(* IEC 61131-3 sources: guidance-for-physical-ai-production-designer-on-aws/source/plan2cell/examples/welding_cell_2_small/plc/trust/robot2/src, 20 files *)

(* ---- E_PlayerState.st ---- *)
(*
 * E_PlayerState
 * States of FB_ProgramPlayer (robot side of the bt2plc zone protocol).
 * Device simulator R2 (robot2), cell welding_cell_2_small. Generated by bt2plc 0.1.0.
 *)

TYPE E_PlayerState :
(
    PS_IDLE         := 0,    (* No program, pose held *)
    PS_NEXT_OP      := 10,   (* Advance to the next op: wStep := k, REQUEST := mask *)
    PS_WAIT_GRANT   := 20,   (* Wait (GRANT AND mask) = mask *)
    PS_DELAY        := 30,   (* Start delay of the op *)
    PS_MOVE         := 40,   (* Trajectory / blind home move *)
    PS_HOLD         := 50,   (* Hold at the end pose *)
    PS_WAIT_RELEASE := 60,   (* REQUEST := 0, wait (GRANT AND mask) = 0 *)
    PS_DONE         := 90,   (* Program finished *)
    PS_ERROR        := 99    (* Program aborted with an error *)
);
END_TYPE

(* ---- E_ProgramState.st ---- *)
(*
 * E_ProgramState
 * VW VASS standard - robot program states.
 * Device simulator R2 (robot2), cell welding_cell_2_small. Generated by bt2plc 0.1.0.
 *)

TYPE E_ProgramState :
(
    PRG_IDLE     := 0,
    PRG_RUNNING  := 1,
    PRG_STOPPED  := 2,
    PRG_PAUSED   := 3,
    PRG_FINISHED := 4,
    PRG_ERROR    := 5
);
END_TYPE

(* ---- E_RobotMode.st ---- *)
(*
 * E_RobotMode
 * VW VASS standard - KUKA KR C4 robot operating modes.
 * Device simulator R2 (robot2), cell welding_cell_2_small. Generated by bt2plc 0.1.0.
 *)

TYPE E_RobotMode :
(
    MODE_UNKNOWN := 0,
    MODE_T1      := 1,       (* Test mode 1 - reduced speed *)
    MODE_T2      := 2,       (* Test mode 2 - programmed speed *)
    MODE_AUT     := 3,       (* Automatic mode *)
    MODE_EXT     := 4        (* External automatic - PLC controlled *)
);
END_TYPE

(* ---- ST_OpDef.st ---- *)
(*
 * ST_OpDef
 * One op of the bt2plc robot program (row of GVL_Program.aOps).
 * Op k plays waypoints GVL_Program.aWp[nFirstWp..nLastWp] under the zone mask dwZoneMask.
 * Blind home op: bBlindHome = TRUE, nFirstWp = nLastWp = 0 (joint move to arHomeDeg over R_HOME_S).
 * Device simulator R2 (robot2), cell welding_cell_2_small. Generated by bt2plc 0.1.0.
 *)

TYPE ST_OpDef :
STRUCT
    sName           : STRING(32);   (* Operation id, e.g. 'W01' *)
    nFirstWp        : INT;          (* First waypoint index in aWp (0 = none) *)
    nLastWp         : INT;          (* Last waypoint index in aWp (0 = none) *)
    dwZoneMask      : DWORD;        (* REQUEST/GRANT bits (zones 0..30, bit 31 = permit) *)
    tDelay          : TIME;         (* Start delay after the grant *)
    tHold           : TIME;         (* Hold time at the end pose *)
    rDelay_s        : REAL;         (* Start delay in s (used by FB_ProgramPlayer) *)
    rHold_s         : REAL;         (* Hold time in s (used by FB_ProgramPlayer) *)
    rVelScale       : REAL;         (* Velocity scale of the trajectory (1.0 = nominal) *)
    bBlindHome      : BOOL;         (* TRUE = blind joint move to the home pose *)
END_STRUCT
END_TYPE

(* ---- ST_PROFIsafe_Trailer.st ---- *)
(*
 * ST_PROFIsafe_Trailer
 * PROFIsafe trailer - 4 bytes appended by the safety layer (status + 3-byte CRC).
 * Device simulator R2 (robot2), cell welding_cell_2_small. Generated by bt2plc 0.1.0.
 *)

TYPE ST_PROFIsafe_Trailer :
STRUCT
    byStatus        : BYTE;                     (* Status/Control byte *)
    abyCRC          : ARRAY[0..2] OF BYTE;      (* 3-byte CRC *)
END_STRUCT
END_TYPE

(* ---- ST_SafeInput.st ---- *)
(*
 * ST_SafeInput
 * PROFIsafe (Slot 1 - FDIO64) safe inputs: robot -> PLC, 8 bytes user data.
 * GSDML: 8x Unsigned8 Input + F_MessageTrailer4Byte.
 * Device simulator R2 (robot2), cell welding_cell_2_small. Generated by bt2plc 0.1.0.
 *)

TYPE ST_SafeInput :
STRUCT
    (* Byte 0: Safe robot status *)
    bSafe_DrivesOK          : BOOL;   (* Bit 0: Safe drives monitoring OK *)
    bSafe_RobotStopped      : BOOL;   (* Bit 1: Robot safely stopped (SOS/SS1) *)
    bSafe_ReducedSpeed      : BOOL;   (* Bit 2: Safe reduced speed active (SLS) *)
    bSafe_AxisMonitoring    : BOOL;   (* Bit 3: Safe axis range monitoring OK *)
    bSafe_ToolOK            : BOOL;   (* Bit 4: Safe tool monitoring OK *)
    bSafe_WorkspaceOK       : BOOL;   (* Bit 5: Safe workspace monitoring OK *)
    bSafe_Reserved06        : BOOL;   (* Bit 6: Reserved *)
    bSafe_Reserved07        : BOOL;   (* Bit 7: Reserved *)

    (* Byte 1: Safe gate/zone status *)
    bSafe_Gate1Closed       : BOOL;   (* Bit 0: Safety gate 1 closed *)
    bSafe_Gate2Closed       : BOOL;   (* Bit 1: Safety gate 2 closed *)
    bSafe_Gate3Closed       : BOOL;   (* Bit 2: Safety gate 3 closed *)
    bSafe_LightCurtainOK    : BOOL;   (* Bit 3: Light curtain free *)
    bSafe_EStopOK           : BOOL;   (* Bit 4: E-Stop not pressed (NC) *)
    bSafe_EnablingDevice    : BOOL;   (* Bit 5: Enabling device pressed (T1/T2) *)
    bSafe_OperatorSafe      : BOOL;   (* Bit 6: Operator protection OK *)
    bSafe_Reserved17        : BOOL;   (* Bit 7: Reserved *)

    (* Byte 2: Extended safe status *)
    bSafe_STO_Active        : BOOL;   (* Bit 0: Safe Torque Off active *)
    bSafe_SS1_Active        : BOOL;   (* Bit 1: Safe Stop 1 active *)
    bSafe_SS2_Active        : BOOL;   (* Bit 2: Safe Stop 2 active *)
    bSafe_SOS_Active        : BOOL;   (* Bit 3: Safe Operating Stop active *)
    bSafe_SLS_Active        : BOOL;   (* Bit 4: Safely-Limited Speed active *)
    bSafe_SLP_Active        : BOOL;   (* Bit 5: Safely-Limited Position active *)
    bSafe_Reserved26        : BOOL;   (* Bit 6: Reserved *)
    bSafe_FaultPresent      : BOOL;   (* Bit 7: Safety fault present *)

    (* Bytes 3-7: Additional safe signals *)
    bySafe_UserInput3       : BYTE;   (* Byte 3: User safe input *)
    bySafe_UserInput4       : BYTE;   (* Byte 4: User safe input *)
    bySafe_UserInput5       : BYTE;   (* Byte 5: User safe input *)
    bySafe_UserInput6       : BYTE;   (* Byte 6: User safe input *)
    bySafe_UserInput7       : BYTE;   (* Byte 7: User safe input *)
END_STRUCT
END_TYPE

(* ---- ST_SafeOutput.st ---- *)
(*
 * ST_SafeOutput
 * PROFIsafe (Slot 1 - FDIO64) safe outputs: PLC -> robot, 8 bytes user data.
 * GSDML: 8x Unsigned8 Output + F_MessageTrailer4Byte.
 * Device simulator R2 (robot2), cell welding_cell_2_small. Generated by bt2plc 0.1.0.
 *)

TYPE ST_SafeOutput :
STRUCT
    (* Byte 0: Safe control from PLC *)
    bSafe_DriveEnable       : BOOL;   (* Bit 0: Enable drives (safe channel) *)
    bSafe_ExternalEStop     : BOOL;   (* Bit 1: External E-Stop request *)
    bSafe_SafeStop1         : BOOL;   (* Bit 2: Request Safe Stop 1 *)
    bSafe_SafeStop2         : BOOL;   (* Bit 3: Request Safe Stop 2 *)
    bSafe_ReducedSpeedReq   : BOOL;   (* Bit 4: Request safe reduced speed *)
    bSafe_GateOverride      : BOOL;   (* Bit 5: Gate override (maintenance) *)
    bSafe_Reserved06        : BOOL;   (* Bit 6: Reserved *)
    bSafe_Reserved07        : BOOL;   (* Bit 7: Reserved *)

    (* Byte 1: Safe zone control *)
    bSafe_Zone1Enable       : BOOL;   (* Bit 0: Enable workspace zone 1 *)
    bSafe_Zone2Enable       : BOOL;   (* Bit 1: Enable workspace zone 2 *)
    bSafe_Zone3Enable       : BOOL;   (* Bit 2: Enable workspace zone 3 *)
    bSafe_Zone4Enable       : BOOL;   (* Bit 3: Enable workspace zone 4 *)
    bSafe_Reserved14        : BOOL;   (* Bit 4: Reserved *)
    bSafe_Reserved15        : BOOL;   (* Bit 5: Reserved *)
    bSafe_Reserved16        : BOOL;   (* Bit 6: Reserved *)
    bSafe_Reserved17        : BOOL;   (* Bit 7: Reserved *)

    (* Bytes 2-7: Additional safe control *)
    bySafe_UserOutput2      : BYTE;   (* Byte 2: User safe output *)
    bySafe_UserOutput3      : BYTE;   (* Byte 3: User safe output *)
    bySafe_UserOutput4      : BYTE;   (* Byte 4: User safe output *)
    bySafe_UserOutput5      : BYTE;   (* Byte 5: User safe output *)
    bySafe_UserOutput6      : BYTE;   (* Byte 6: User safe output *)
    bySafe_UserOutput7      : BYTE;   (* Byte 7: User safe output *)
END_STRUCT
END_TYPE

(* ---- ST_VASS_ControlWord.st ---- *)
(*
 * ST_VASS_ControlWord
 * VASS PLC control word - output bytes 0-1 (PLC -> robot), Slot 2 DIO256.
 * Device simulator R2 (robot2), cell welding_cell_2_small. Generated by bt2plc 0.1.0.
 *)

TYPE ST_VASS_ControlWord :
STRUCT
    (* Byte 0 *)
    bDrivesOn           : BOOL;   (* Bit 0: Enable drives *)
    bProgStart          : BOOL;   (* Bit 1: Start program *)
    bProgStop           : BOOL;   (* Bit 2: Stop program *)
    bProgCancel         : BOOL;   (* Bit 3: Cancel program *)
    bModeRequest        : BOOL;   (* Bit 4: Request EXT mode *)
    bReset              : BOOL;   (* Bit 5: Reset error *)
    bHomeRequest        : BOOL;   (* Bit 6: Move to home *)
    bConfirm            : BOOL;   (* Bit 7: Confirm/acknowledge *)

    (* Byte 1 *)
    bJobRequest         : BOOL;   (* Bit 8: New job request *)
    bGripperOpen        : BOOL;   (* Bit 9: Open gripper *)
    bGripperClose       : BOOL;   (* Bit 10: Close gripper *)
    bPeriphRelease      : BOOL;   (* Bit 11: Release peripheral *)
    bSpeedOverride      : BOOL;   (* Bit 12: Apply speed override *)
    bReserved13         : BOOL;   (* Bit 13: Reserved *)
    bReserved14         : BOOL;   (* Bit 14: Reserved *)
    bReserved15         : BOOL;   (* Bit 15: Reserved *)
END_STRUCT
END_TYPE

(* ---- ST_VASS_InputTelegram.st ---- *)
(*
 * ST_VASS_InputTelegram
 * Full VASS input telegram - 32 bytes (robot -> PLC), Slot 2 DIO256 inputs.
 * bt2plc use: bytes 4-5 wCurrentStep = op index (GVL_Program.STEP_BYTE),
 *             bytes 16-27 joint angles A1..A6 (FB_JointAngleEncoder),
 *             bytes 28-31 zone REQUEST DWORD LE (GVL_Program.REQ_BYTE).
 * Device simulator R2 (robot2), cell welding_cell_2_small. Generated by bt2plc 0.1.0.
 *)

TYPE ST_VASS_InputTelegram :
STRUCT
    stStatusWord        : ST_VASS_StatusWord;     (* Bytes 0-1:   Status word *)
    wActiveJobNr        : WORD;                   (* Bytes 2-3:   Active job number *)
    wCurrentStep        : WORD;                   (* Bytes 4-5:   Current program step *)
    wSpeedActual        : WORD;                   (* Bytes 6-7:   Actual speed % *)
    wActiveToolNr       : WORD;                   (* Bytes 8-9:   Active tool number *)
    wErrorCode          : WORD;                   (* Bytes 10-11: Active error code *)
    wWarningCode        : WORD;                   (* Bytes 12-13: Active warning code *)
    wPositionX          : INT;                    (* Bytes 14-15: Position X (0.1mm) *)
    wPositionY          : INT;                    (* Bytes 16-17: Position Y (0.1mm) *)
    wPositionZ          : INT;                    (* Bytes 18-19: Position Z (0.1mm) *)
    wUserWord10         : WORD;                   (* Bytes 20-21: User data *)
    wUserWord11         : WORD;                   (* Bytes 22-23: User data *)
    wUserWord12         : WORD;                   (* Bytes 24-25: User data *)
    wUserWord13         : WORD;                   (* Bytes 26-27: User data *)
    wUserWord14         : WORD;                   (* Bytes 28-29: User data *)
    wUserWord15         : WORD;                   (* Bytes 30-31: User data *)
END_STRUCT
END_TYPE

(* ---- ST_VASS_OutputTelegram.st ---- *)
(*
 * ST_VASS_OutputTelegram
 * Full VASS output telegram - 32 bytes (PLC -> robot), Slot 2 DIO256 outputs.
 * bt2plc use: bytes 4-5 PLAN_ID WORD LE during a production job (GVL_Program.PLAN_ID_BYTE),
 *             bytes 12-15 zone GRANT DWORD LE (GVL_Program.GRANT_BYTE).
 * Device simulator R2 (robot2), cell welding_cell_2_small. Generated by bt2plc 0.1.0.
 *)

TYPE ST_VASS_OutputTelegram :
STRUCT
    stControlWord       : ST_VASS_ControlWord;    (* Bytes 0-1:   Control word *)
    wJobNr              : WORD;                   (* Bytes 2-3:   Requested job number *)
    wParameter1         : WORD;                   (* Bytes 4-5:   Parameter 1 *)
    wParameter2         : WORD;                   (* Bytes 6-7:   Parameter 2 *)
    wSpeedOverride      : WORD;                   (* Bytes 8-9:   Speed override % *)
    wToolRequest        : WORD;                   (* Bytes 10-11: Tool change request *)
    wUserWord6          : WORD;                   (* Bytes 12-13: User command data *)
    wUserWord7          : WORD;                   (* Bytes 14-15: User command data *)
    wUserWord8          : WORD;                   (* Bytes 16-17: User command data *)
    wUserWord9          : WORD;                   (* Bytes 18-19: User command data *)
    wUserWord10         : WORD;                   (* Bytes 20-21: User command data *)
    wUserWord11         : WORD;                   (* Bytes 22-23: User command data *)
    wUserWord12         : WORD;                   (* Bytes 24-25: User command data *)
    wUserWord13         : WORD;                   (* Bytes 26-27: User command data *)
    wUserWord14         : WORD;                   (* Bytes 28-29: User command data *)
    wUserWord15         : WORD;                   (* Bytes 30-31: User command data *)
END_STRUCT
END_TYPE

(* ---- ST_VASS_StatusWord.st ---- *)
(*
 * ST_VASS_StatusWord
 * VASS robot status word - input bytes 0-1 (robot -> PLC), Slot 2 DIO256.
 * Device simulator R2 (robot2), cell welding_cell_2_small. Generated by bt2plc 0.1.0.
 *)

TYPE ST_VASS_StatusWord :
STRUCT
    (* Byte 0 *)
    bDrivesPowered      : BOOL;   (* Bit 0: Drives are powered on *)
    bProgRunning        : BOOL;   (* Bit 1: Program is running *)
    bAtHome             : BOOL;   (* Bit 2: Robot at home position *)
    bInPosition         : BOOL;   (* Bit 3: Robot in target position *)
    bModeExt            : BOOL;   (* Bit 4: External automatic mode active *)
    bReady              : BOOL;   (* Bit 5: Robot ready for command *)
    bError              : BOOL;   (* Bit 6: Error present *)
    bWarning            : BOOL;   (* Bit 7: Warning present *)

    (* Byte 1 *)
    bSafetyGateOK       : BOOL;   (* Bit 8: Safety gate closed *)
    bEStopNotActive     : BOOL;   (* Bit 9: E-Stop NOT active (NC logic) *)
    bProgFinished       : BOOL;   (* Bit 10: Program/job finished *)
    bJobAcknowledge     : BOOL;   (* Bit 11: Job number acknowledged *)
    bToolActive         : BOOL;   (* Bit 12: Tool/gripper active *)
    bPartPresent        : BOOL;   (* Bit 13: Part present in gripper *)
    bPeriphReady        : BOOL;   (* Bit 14: Peripheral devices ready *)
    bMaintRequired      : BOOL;   (* Bit 15: Maintenance required *)
END_STRUCT
END_TYPE

(* ---- ST_Waypoint.st ---- *)
(*
 * ST_Waypoint
 * One trajectory waypoint (row of GVL_Program.aWp). Flat fields for portability.
 * rT = seconds from op start; angles in degrees (KUKA A1..A6 after joint sign/offset mapping).
 * Device simulator R2 (robot2), cell welding_cell_2_small. Generated by bt2plc 0.1.0.
 *)

TYPE ST_Waypoint :
STRUCT
    rT              : REAL;         (* Time from op start (s) *)
    rA1             : REAL;         (* Axis 1 (deg) *)
    rA2             : REAL;         (* Axis 2 (deg) *)
    rA3             : REAL;         (* Axis 3 (deg) *)
    rA4             : REAL;         (* Axis 4 (deg) *)
    rA5             : REAL;         (* Axis 5 (deg) *)
    rA6             : REAL;         (* Axis 6 (deg) *)
END_STRUCT
END_TYPE

(* ---- GVL_DeviceParams.st ---- *)
NAMESPACE GVL_DeviceParams
(*
 * GVL_DeviceParams
 * PROFINET device identity parameters.
 * Device simulator R2 (robot2, station kuka-robi2), cell welding_cell_2_small. Generated by bt2plc 0.1.0.
 *
 * These parameters configure how the CODESYS PROFINET Device presents itself
 * on the network. They MUST match what the Siemens PLC expects (from the GSDML).
 *
 * In CODESYS, these are typically set via:
 *   1. The "PROFINET Device IEC Objects" tab in the device editor
 *   2. Or programmatically by writing to the device parameter structure
 *
 * The CODESYS PROFINET Device stack reads these at startup and uses them
 * in DCP responses and during the PROFINET connection establishment.
 *
 * IMPORTANT: The default CODESYS values (VendorId=0x02CC, DeviceId=0x1017)
 * will NOT work with the Siemens PLC that expects KUKA (0x019B / 0x0301).
 * You MUST override them.
 *)

{attribute 'qualified_only'}
VAR_GLOBAL
    (* === KUKA VKRCnexxt Device Identity === *)
    (* These values come from GSDML-V2.25-KUKA-Roboter-GmbH-VKR C4-Device-V1.0 *)

    VENDOR_ID           : UINT        := 16#019B;                 (* KUKA Roboter GmbH *)
    DEVICE_ID           : UINT        := 16#0301;                 (* VKR C4 Device *)
    STATION_TYPE        : STRING(240) := 'KUKA VKR C4';           (* Station type string *)
    DEVICE_TYPE         : STRING(28)  := 'KUKA VKR C4';           (* Device type string *)
    ORDER_ID            : STRING(20)  := 'KUKA VKRC nexxt';       (* Order number *)
    HW_REVISION         : UINT        := 1;                       (* Hardware revision *)
    SW_REV_PREFIX       : USINT       := 16#56;                   (* 'V' in ASCII *)
    SW_REV_MAJOR        : UINT        := 8;                       (* V8.x *)
    SW_REV_MINOR        : UINT        := 2;                       (* x.2 *)
    SW_REV_PATCH        : UINT        := 0;                       (* x.x.0 *)

    (* === Module Identification Numbers (from GSDML) === *)
    MODULE_IDENT_DAP    : DWORD       := DWORD#16#00000301;       (* DAP - Slot 0 *)
    MODULE_IDENT_FDIO64 : DWORD       := DWORD#16#0000008F;       (* PROFIsafe - Slot 1 *)
    MODULE_IDENT_DIO256 : DWORD       := DWORD#16#00001000;       (* VASS telegram - Slot 2 *)
    SUBMODULE_IDENT     : DWORD       := DWORD#16#00000001;       (* Submodule ident (all slots) *)

    (* === PROFIsafe Parameters (Slot 1) === *)
    (* These must match the F-parameter record in the PLC safety configuration *)
    F_SIL_LEVEL         : UINT        := 3;                       (* SIL 3 *)
    F_CRC_LENGTH        : UINT        := 3;                       (* 3-byte CRC *)
    F_WD_TIME_DEFAULT   : UINT        := 500;                     (* Watchdog 500ms *)
    F_BLOCK_ID          : UINT        := 0;                       (* Block ID *)
    F_PAR_CRC_DEFAULT   : UINT        := 16#FF59;                 (* Default F_Par_CRC = 65369 *)
END_VAR
END_NAMESPACE

(* ---- GVL_IO.st ---- *)
NAMESPACE GVL_IO
(*
 * GVL_IO
 * Global variable list for the PROFINET device I/O mapping.
 * Device simulator R2 (robot2, station kuka-robi2), cell welding_cell_2_small. Generated by bt2plc 0.1.0.
 *
 * These variables are mapped to the PROFINET device modules via the I/O Mapping tab.
 * Do NOT use AT addresses - the mapping is done in the device configuration.
 * Only PLC_PRG accesses this GVL: it copies the commands into local images and writes
 * the robot status back as a whole array / as scalars (the FBs never touch GVL_IO).
 *
 * Module mapping (set in I/O Mapping tab of each module):
 *   SafeIO_FDIO64 (Slot 1):
 *     "8 safe digital inputs" channels  -> GVL_IO.bySafeIn0..bySafeIn7
 *     "8 safe digital outputs" channels -> GVL_IO.bySafeOut0..bySafeOut7
 *
 *   VASS_DIO256 (Slot 2):
 *     Input channel  -> GVL_IO.aVassInputData
 *     Output channel -> GVL_IO.aVassOutputData
 *)

{attribute 'qualified_only'}
VAR_GLOBAL
    (* ========================================================================
       SLOT 1 - PROFIsafe FDIO64 Module
       8 individual USINT/BYTE channels per direction
       Map each one to the corresponding "8 safe digital inputs/outputs" row
       ======================================================================== *)

    (* Safe Inputs: Robot -> PLC (mapped to "8 safe digital inputs" channels) *)
    bySafeIn0       : BYTE;     (* Safe input byte 0: Drive status *)
    bySafeIn1       : BYTE;     (* Safe input byte 1: Gate/protection *)
    bySafeIn2       : BYTE;     (* Safe input byte 2: STO/SS1/SS2/SOS/SLS *)
    bySafeIn3       : BYTE;     (* Safe input byte 3: User *)
    bySafeIn4       : BYTE;     (* Safe input byte 4: User *)
    bySafeIn5       : BYTE;     (* Safe input byte 5: User *)
    bySafeIn6       : BYTE;     (* Safe input byte 6: User *)
    bySafeIn7       : BYTE;     (* Safe input byte 7: User *)

    (* Safe Outputs: PLC -> Robot (mapped to "8 safe digital outputs" channels) *)
    bySafeOut0      : BYTE;     (* Safe output byte 0: Drive enable, E-Stop, SS1/SS2 *)
    bySafeOut1      : BYTE;     (* Safe output byte 1: Zone enables *)
    bySafeOut2      : BYTE;     (* Safe output byte 2: User *)
    bySafeOut3      : BYTE;     (* Safe output byte 3: User *)
    bySafeOut4      : BYTE;     (* Safe output byte 4: User *)
    bySafeOut5      : BYTE;     (* Safe output byte 5: User *)
    bySafeOut6      : BYTE;     (* Safe output byte 6: User *)
    bySafeOut7      : BYTE;     (* Safe output byte 7: User *)

    (* ========================================================================
       SLOT 2 - DIO256 VASS Telegram
       32 bytes per direction as arrays
       ======================================================================== *)

    (* VASS Inputs: Robot -> PLC (32 bytes) *)
    aVassInputData      : ARRAY[0..31] OF BYTE;

    (* VASS Outputs: PLC -> Robot (32 bytes) *)
    aVassOutputData     : ARRAY[0..31] OF BYTE;
END_VAR
END_NAMESPACE

(* ---- GVL_Program.st ---- *)
NAMESPACE GVL_Program
(*
 * GVL_Program - generated by bt2plc 0.1.0 - DO NOT EDIT
 * Robot program of robot2 (R2) for plan bt_1790934549_welding_cell_2_small (cell welding_cell_2_small)
 * Angles in degrees (KUKA A1..A6 after joint sign/offset), times in seconds from op start.
 *)
{attribute 'qualified_only'}
VAR_GLOBAL
    (* ========================================================================
       IDENTITY / PROTOCOL
       ======================================================================== *)
    ROBOT_TAG               : STRING(16) := 'R2';
    ROBOT_NS                : STRING(32) := 'robot2';
    ROBOT_INDEX             : WORD := WORD#2;
    PLAN_ID                 : WORD := WORD#16#F77E;             (* must match the head PLC *)
    PROD_FOLGE              : WORD := WORD#11;
    HOME_FOLGE              : WORD := WORD#125;
    JOB_NUMBER_BYTE         : BOOL := FALSE;
    STEP_BYTE               : INT := 4;
    REQ_BYTE                : INT := 28;
    GRANT_BYTE              : INT := 12;
    PLAN_ID_BYTE            : INT := 4;
    R_TASK_S                : REAL := 0.0200;                   (* device MainTask interval *)
    R_HOME_S                : REAL := 7.0000;                   (* blind home duration *)
    R_AT_HOME_TOL_DEG       : REAL := 0.5000;
    R_START_TOL_DEG         : REAL := 1.0000;
    ERR_UNKNOWN_FOLGE       : WORD := WORD#16#0101;
    ERR_PLAN_MISMATCH       : WORD := WORD#16#0103;
    WARN_START_DEVIATION    : WORD := WORD#16#0201;

    (* ========================================================================
       PROGRAM
       ======================================================================== *)
    N_OPS                   : INT := 10;
    N_WP                    : INT := 263;
    arHomeDeg               : ARRAY[1..6] OF REAL := [0.0000, -90.0000, 90.0000, 0.0000, 0.0000, 0.0000];
    aOps                    : ARRAY[1..10] OF ST_OpDef := [
        (sName := 'W13', nFirstWp := 1, nLastWp := 41, dwZoneMask := DWORD#16#00000002, tDelay := T#0MS, tHold := T#500MS, rDelay_s := 0.0000, rHold_s := 0.5000, rVelScale := 1.0000, bBlindHome := FALSE),    (* #1 W13 (weld) *)
        (sName := 'W15', nFirstWp := 42, nLastWp := 77, dwZoneMask := DWORD#16#00000001, tDelay := T#0MS, tHold := T#500MS, rDelay_s := 0.0000, rHold_s := 0.5000, rVelScale := 1.0000, bBlindHome := FALSE),    (* #2 W15 (weld) *)
        (sName := 'W14', nFirstWp := 78, nLastWp := 100, dwZoneMask := DWORD#16#00000002, tDelay := T#0MS, tHold := T#500MS, rDelay_s := 0.0000, rHold_s := 0.5000, rVelScale := 1.0000, bBlindHome := FALSE),    (* #3 W14 (weld) *)
        (sName := 'W10', nFirstWp := 101, nLastWp := 124, dwZoneMask := DWORD#16#00000001, tDelay := T#0MS, tHold := T#500MS, rDelay_s := 0.0000, rHold_s := 0.5000, rVelScale := 1.0000, bBlindHome := FALSE),    (* #4 W10 (weld) *)
        (sName := 'W11', nFirstWp := 125, nLastWp := 148, dwZoneMask := DWORD#16#00000002, tDelay := T#0MS, tHold := T#500MS, rDelay_s := 0.0000, rHold_s := 0.5000, rVelScale := 1.0000, bBlindHome := FALSE),    (* #5 W11 (weld) *)
        (sName := 'W12', nFirstWp := 149, nLastWp := 171, dwZoneMask := DWORD#16#00000001, tDelay := T#0MS, tHold := T#500MS, rDelay_s := 0.0000, rHold_s := 0.5000, rVelScale := 1.0000, bBlindHome := FALSE),    (* #6 W12 (weld) *)
        (sName := 'W09', nFirstWp := 172, nLastWp := 186, dwZoneMask := DWORD#16#00000001, tDelay := T#0MS, tHold := T#500MS, rDelay_s := 0.0000, rHold_s := 0.5000, rVelScale := 1.0000, bBlindHome := FALSE),    (* #7 W09 (weld) *)
        (sName := 'W08', nFirstWp := 187, nLastWp := 208, dwZoneMask := DWORD#16#00000000, tDelay := T#0MS, tHold := T#500MS, rDelay_s := 0.0000, rHold_s := 0.5000, rVelScale := 1.0000, bBlindHome := FALSE),    (* #8 W08 (weld) *)
        (sName := 'W07', nFirstWp := 209, nLastWp := 231, dwZoneMask := DWORD#16#00000002, tDelay := T#0MS, tHold := T#500MS, rDelay_s := 0.0000, rHold_s := 0.5000, rVelScale := 1.0000, bBlindHome := FALSE),    (* #9 W07 (weld) *)
        (sName := 'HOME', nFirstWp := 232, nLastWp := 263, dwZoneMask := DWORD#16#00000000, tDelay := T#0MS, tHold := T#0MS, rDelay_s := 0.0000, rHold_s := 0.0000, rVelScale := 1.0000, bBlindHome := FALSE)    (* #10 HOME (home) *)
    ];
    aWp                     : ARRAY[1..263] OF ST_Waypoint := [
        (* op 1 W13 - traj_robot2_W13 *)
        (rT := 0.0000, rA1 := 0.0000, rA2 := -90.0000, rA3 := 90.0000, rA4 := 0.0000, rA5 := 0.0000, rA6 := 0.0000),
        (rT := 0.2730, rA1 := 0.3035, rA2 := -89.9642, rA3 := 90.0888, rA4 := -0.1637, rA5 := 0.2135, rA6 := -0.1916),
        (rT := 0.5457, rA1 := 1.1862, rA2 := -89.8601, rA3 := 90.3471, rA4 := -0.6399, rA5 := 0.8344, rA6 := -0.7490),
        (rT := 0.8187, rA1 := 2.6069, rA2 := -89.6924, rA3 := 90.7628, rA4 := -1.4062, rA5 := 1.8337, rA6 := -1.6461),
        (rT := 1.0913, rA1 := 4.5242, rA2 := -89.4662, rA3 := 91.3239, rA4 := -2.4404, rA5 := 3.1824, rA6 := -2.8567),
        (rT := 1.3643, rA1 := 6.8967, rA2 := -89.1864, rA3 := 92.0181, rA4 := -3.7201, rA5 := 4.8512, rA6 := -4.3548),
        (rT := 1.6373, rA1 := 9.6830, rA2 := -88.8576, rA3 := 92.8334, rA4 := -5.2230, rA5 := 6.8110, rA6 := -6.1141),
        (rT := 1.9100, rA1 := 12.8416, rA2 := -88.4850, rA3 := 93.7577, rA4 := -6.9268, rA5 := 9.0329, rA6 := -8.1086),
        (rT := 2.1830, rA1 := 16.3314, rA2 := -88.0733, rA3 := 94.7788, rA4 := -8.8092, rA5 := 11.4875, rA6 := -10.3121),
        (rT := 2.4557, rA1 := 20.1107, rA2 := -87.6274, rA3 := 95.8848, rA4 := -10.8478, rA5 := 14.1460, rA6 := -12.6985),
        (rT := 2.7287, rA1 := 24.1384, rA2 := -87.1522, rA3 := 97.0633, rA4 := -13.0204, rA5 := 16.9790, rA6 := -15.2417),
        (rT := 3.0017, rA1 := 28.3730, rA2 := -86.6527, rA3 := 98.3024, rA4 := -15.3045, rA5 := 19.9577, rA6 := -17.9155),
        (rT := 3.2743, rA1 := 32.7731, rA2 := -86.1336, rA3 := 99.5900, rA4 := -17.6779, rA5 := 23.0527, rA6 := -20.6938),
        (rT := 3.5473, rA1 := 37.2973, rA2 := -85.5998, rA3 := 100.9138, rA4 := -20.1183, rA5 := 26.2351, rA6 := -23.5505),
        (rT := 3.8203, rA1 := 41.9043, rA2 := -85.0563, rA3 := 102.2619, rA4 := -22.6034, rA5 := 29.4756, rA6 := -26.4595),
        (rT := 4.0930, rA1 := 46.5527, rA2 := -84.5079, rA3 := 103.6221, rA4 := -25.1107, rA5 := 32.7453, rA6 := -29.3946),
        (rT := 4.3660, rA1 := 51.2010, rA2 := -83.9595, rA3 := 104.9823, rA4 := -27.6181, rA5 := 36.0150, rA6 := -32.3297),
        (rT := 4.6387, rA1 := 55.8080, rA2 := -83.4160, rA3 := 106.3304, rA4 := -30.1031, rA5 := 39.2556, rA6 := -35.2387),
        (rT := 4.9117, rA1 := 60.3322, rA2 := -82.8822, rA3 := 107.6543, rA4 := -32.5435, rA5 := 42.4379, rA6 := -38.0954),
        (rT := 5.1847, rA1 := 64.7323, rA2 := -82.3631, rA3 := 108.9418, rA4 := -34.9169, rA5 := 45.5329, rA6 := -40.8738),
        (rT := 5.4573, rA1 := 68.9669, rA2 := -81.8635, rA3 := 110.1809, rA4 := -37.2011, rA5 := 48.5116, rA6 := -43.5476),
        (rT := 5.7303, rA1 := 72.9946, rA2 := -81.3884, rA3 := 111.3595, rA4 := -39.3736, rA5 := 51.3446, rA6 := -46.0908),
        (rT := 6.0030, rA1 := 76.7740, rA2 := -80.9425, rA3 := 112.4654, rA4 := -41.4122, rA5 := 54.0031, rA6 := -48.4772),
        (rT := 6.2760, rA1 := 80.2637, rA2 := -80.5308, rA3 := 113.4866, rA4 := -43.2946, rA5 := 56.4578, rA6 := -50.6807),
        (rT := 6.5490, rA1 := 83.4224, rA2 := -80.1581, rA3 := 114.4108, rA4 := -44.9984, rA5 := 58.6796, rA6 := -52.6752),
        (rT := 6.8217, rA1 := 86.2086, rA2 := -79.8294, rA3 := 115.2262, rA4 := -46.5013, rA5 := 60.6394, rA6 := -54.4345),
        (rT := 7.0947, rA1 := 88.5811, rA2 := -79.5495, rA3 := 115.9204, rA4 := -47.7810, rA5 := 62.3082, rA6 := -55.9325),
        (rT := 7.3673, rA1 := 90.4984, rA2 := -79.3233, rA3 := 116.4814, rA4 := -48.8152, rA5 := 63.6569, rA6 := -57.1431),
        (rT := 7.6403, rA1 := 91.9191, rA2 := -79.1557, rA3 := 116.8971, rA4 := -49.5816, rA5 := 64.6562, rA6 := -58.0402),
        (rT := 7.9133, rA1 := 92.8019, rA2 := -79.0516, rA3 := 117.1554, rA4 := -50.0578, rA5 := 65.2772, rA6 := -58.5976),
        (rT := 8.1860, rA1 := 93.1053, rA2 := -79.0158, rA3 := 117.2442, rA4 := -50.2214, rA5 := 65.4906, rA6 := -58.7892),
        (rT := 8.2860, rA1 := 93.1054, rA2 := -78.5375, rA3 := 117.5788, rA4 := -50.4217, rA5 := 65.3570, rA6 := -58.5702),
        (rT := 8.3860, rA1 := 93.1056, rA2 := -77.8336, rA3 := 118.0660, rA4 := -50.7525, rA5 := 65.1056, rA6 := -58.1705),
        (rT := 8.4860, rA1 := 93.1056, rA2 := -77.4884, rA3 := 118.2931, rA4 := -51.0112, rA5 := 64.8431, rA6 := -57.7771),
        (rT := 8.5860, rA1 := 93.1055, rA2 := -77.2114, rA3 := 118.4657, rA4 := -51.2652, rA5 := 64.5476, rA6 := -57.3432),
        (rT := 8.6860, rA1 := 93.1055, rA2 := -76.8948, rA3 := 118.6607, rA4 := -51.5186, rA5 := 64.2245, rA6 := -56.8729),
        (rT := 8.7860, rA1 := 93.1055, rA2 := -76.5752, rA3 := 118.8523, rA4 := -51.7590, rA5 := 63.8986, rA6 := -56.4005),
        (rT := 8.8860, rA1 := 93.1055, rA2 := -76.2532, rA3 := 119.0400, rA4 := -51.9657, rA5 := 63.6083, rA6 := -55.9794),
        (rT := 8.9860, rA1 := 93.1055, rA2 := -75.9277, rA3 := 119.2244, rA4 := -52.1675, rA5 := 63.3171, rA6 := -55.5556),
        (rT := 9.0860, rA1 := 93.1055, rA2 := -75.5136, rA3 := 119.4506, rA4 := -52.4491, rA5 := 62.9118, rA6 := -54.9605),
        (rT := 9.1860, rA1 := 93.1055, rA2 := -75.2634, rA3 := 119.5852, rA4 := -52.6226, rA5 := 62.6611, rA6 := -54.5914),
        (* op 2 W15 - traj_robot2_W15 *)
        (rT := 0.0000, rA1 := 93.1055, rA2 := -75.2634, rA3 := 119.5852, rA4 := -52.6226, rA5 := 62.6611, rA6 := -54.5914),
        (rT := 0.2770, rA1 := 93.0446, rA2 := -75.3085, rA3 := 119.5681, rA4 := -52.1640, rA5 := 62.7161, rA6 := -54.8912),
        (rT := 0.5540, rA1 := 92.8686, rA2 := -75.4391, rA3 := 119.5185, rA4 := -50.8385, rA5 := 62.8751, rA6 := -55.7578),
        (rT := 0.8310, rA1 := 92.5874, rA2 := -75.6476, rA3 := 119.4393, rA4 := -48.7214, rA5 := 63.1291, rA6 := -57.1419),
        (rT := 1.1080, rA1 := 92.2111, rA2 := -75.9266, rA3 := 119.3333, rA4 := -45.8882, rA5 := 63.4690, rA6 := -58.9942),
        (rT := 1.3850, rA1 := 91.7498, rA2 := -76.2688, rA3 := 119.2033, rA4 := -42.4142, rA5 := 63.8858, rA6 := -61.2654),
        (rT := 1.6620, rA1 := 91.2133, rA2 := -76.6667, rA3 := 119.0521, rA4 := -38.3748, rA5 := 64.3703, rA6 := -63.9062),
        (rT := 1.9390, rA1 := 90.6118, rA2 := -77.1128, rA3 := 118.8827, rA4 := -33.8454, rA5 := 64.9137, rA6 := -66.8675),
        (rT := 2.2160, rA1 := 89.9552, rA2 := -77.5997, rA3 := 118.6977, rA4 := -28.9013, rA5 := 65.5068, rA6 := -70.0997),
        (rT := 2.4930, rA1 := 89.2535, rA2 := -78.1201, rA3 := 118.5000, rA4 := -23.6181, rA5 := 66.1406, rA6 := -73.5538),
        (rT := 2.7700, rA1 := 88.5168, rA2 := -78.6664, rA3 := 118.2925, rA4 := -18.0710, rA5 := 66.8061, rA6 := -77.1803),
        (rT := 3.0470, rA1 := 87.7551, rA2 := -79.2313, rA3 := 118.0779, rA4 := -12.3354, rA5 := 67.4942, rA6 := -80.9301),
        (rT := 3.3240, rA1 := 86.9784, rA2 := -79.8073, rA3 := 117.8590, rA4 := -6.4867, rA5 := 68.1958, rA6 := -84.7538),
        (rT := 3.6010, rA1 := 86.1966, rA2 := -80.3871, rA3 := 117.6388, rA4 := -0.6004, rA5 := 68.9020, rA6 := -88.6021),
        (rT := 3.8780, rA1 := 85.4199, rA2 := -80.9631, rA3 := 117.4200, rA4 := 5.2483, rA5 := 69.6036, rA6 := -92.4258),
        (rT := 4.1550, rA1 := 84.6581, rA2 := -81.5280, rA3 := 117.2054, rA4 := 10.9839, rA5 := 70.2917, rA6 := -96.1756),
        (rT := 4.4320, rA1 := 83.9214, rA2 := -82.0744, rA3 := 116.9978, rA4 := 16.5310, rA5 := 70.9571, rA6 := -99.8021),
        (rT := 4.7090, rA1 := 83.2198, rA2 := -82.5947, rA3 := 116.8002, rA4 := 21.8142, rA5 := 71.5909, rA6 := -103.2562),
        (rT := 4.9860, rA1 := 82.5632, rA2 := -83.0817, rA3 := 116.6152, rA4 := 26.7583, rA5 := 72.1840, rA6 := -106.4884),
        (rT := 5.2630, rA1 := 81.9617, rA2 := -83.5278, rA3 := 116.4457, rA4 := 31.2877, rA5 := 72.7274, rA6 := -109.4496),
        (rT := 5.5400, rA1 := 81.4252, rA2 := -83.9256, rA3 := 116.2946, rA4 := 35.3271, rA5 := 73.2120, rA6 := -112.0905),
        (rT := 5.8170, rA1 := 80.9638, rA2 := -84.2678, rA3 := 116.1646, rA4 := 38.8011, rA5 := 73.6288, rA6 := -114.3617),
        (rT := 6.0940, rA1 := 80.5876, rA2 := -84.5468, rA3 := 116.0586, rA4 := 41.6343, rA5 := 73.9686, rA6 := -116.2140),
        (rT := 6.3710, rA1 := 80.3064, rA2 := -84.7554, rA3 := 115.9794, rA4 := 43.7514, rA5 := 74.2226, rA6 := -117.5981),
        (rT := 6.6480, rA1 := 80.1303, rA2 := -84.8859, rA3 := 115.9298, rA4 := 45.0769, rA5 := 74.3816, rA6 := -118.4647),
        (rT := 6.9250, rA1 := 80.0694, rA2 := -84.9311, rA3 := 115.9126, rA4 := 45.5355, rA5 := 74.4367, rA6 := -118.7645),
        (rT := 7.0250, rA1 := 80.0693, rA2 := -84.5291, rA3 := 116.3283, rA4 := 45.7971, rA5 := 74.2601, rA6 := -119.1812),
        (rT := 7.1250, rA1 := 80.0690, rA2 := -83.9370, rA3 := 116.9342, rA4 := 46.1788, rA5 := 73.9509, rA6 := -119.8289),
        (rT := 7.2250, rA1 := 80.0690, rA2 := -83.6457, rA3 := 117.2174, rA4 := 46.3591, rA5 := 73.6768, rA6 := -120.2334),
        (rT := 7.3250, rA1 := 80.0690, rA2 := -83.4107, rA3 := 117.4340, rA4 := 46.4966, rA5 := 73.3758, rA6 := -120.6123),
        (rT := 7.4250, rA1 := 80.0690, rA2 := -83.1411, rA3 := 117.6800, rA4 := 46.6500, rA5 := 73.0334, rA6 := -121.0389),
        (rT := 7.5250, rA1 := 80.0690, rA2 := -82.8676, rA3 := 117.9231, rA4 := 46.7976, rA5 := 72.6753, rA6 := -121.4706),
        (rT := 7.6250, rA1 := 80.0690, rA2 := -82.5907, rA3 := 118.1628, rA4 := 46.9371, rA5 := 72.3209, rA6 := -121.8897),
        (rT := 7.7250, rA1 := 80.0690, rA2 := -82.3101, rA3 := 118.3993, rA4 := 47.0693, rA5 := 71.9737, rA6 := -122.2947),
        (rT := 7.8250, rA1 := 80.0690, rA2 := -81.9537, rA3 := 118.6895, rA4 := 47.2230, rA5 := 71.5682, rA6 := -122.7657),
        (rT := 7.9250, rA1 := 80.0690, rA2 := -81.7384, rA3 := 118.8624, rA4 := 47.3124, rA5 := 71.3307, rA6 := -123.0405),
        (* op 3 W14 - traj_robot2_W14 *)
        (rT := 0.0000, rA1 := 80.0690, rA2 := -81.7384, rA3 := 118.8624, rA4 := 47.3124, rA5 := 71.3307, rA6 := -123.0405),
        (rT := 0.2687, rA1 := 80.1323, rA2 := -81.6821, rA3 := 118.7100, rA4 := 46.4005, rA5 := 71.0643, rA6 := -122.5345),
        (rT := 0.5373, rA1 := 80.3070, rA2 := -81.5266, rA3 := 118.2888, rA4 := 43.8793, rA5 := 70.3279, rA6 := -121.1355),
        (rT := 0.8060, rA1 := 80.5710, rA2 := -81.2918, rA3 := 117.6524, rA4 := 40.0706, rA5 := 69.2153, rA6 := -119.0220),
        (rT := 1.0747, rA1 := 80.9020, rA2 := -80.9973, rA3 := 116.8546, rA4 := 35.2964, rA5 := 67.8207, rA6 := -116.3728),
        (rT := 1.3433, rA1 := 81.2775, rA2 := -80.6632, rA3 := 115.9494, rA4 := 29.8784, rA5 := 66.2380, rA6 := -113.3663),
        (rT := 1.6120, rA1 := 81.6754, rA2 := -80.3092, rA3 := 114.9903, rA4 := 24.1386, rA5 := 64.5614, rA6 := -110.1813),
        (rT := 1.8807, rA1 := 82.0732, rA2 := -79.9553, rA3 := 114.0312, rA4 := 18.3988, rA5 := 62.8847, rA6 := -106.9963),
        (rT := 2.1493, rA1 := 82.4488, rA2 := -79.6211, rA3 := 113.1260, rA4 := 12.9808, rA5 := 61.3021, rA6 := -103.9898),
        (rT := 2.4180, rA1 := 82.7797, rA2 := -79.3267, rA3 := 112.3282, rA4 := 8.2066, rA5 := 59.9075, rA6 := -101.3406),
        (rT := 2.6867, rA1 := 83.0437, rA2 := -79.0918, rA3 := 111.6919, rA4 := 4.3979, rA5 := 58.7949, rA6 := -99.2271),
        (rT := 2.9553, rA1 := 83.2185, rA2 := -78.9363, rA3 := 111.2706, rA4 := 1.8767, rA5 := 58.0584, rA6 := -97.8281),
        (rT := 3.2243, rA1 := 83.2817, rA2 := -78.8801, rA3 := 111.1182, rA4 := 0.9647, rA5 := 57.7920, rA6 := -97.3221),
        (rT := 3.3243, rA1 := 83.2819, rA2 := -78.5511, rA3 := 111.4303, rA4 := 0.7191, rA5 := 57.4498, rA6 := -97.1693),
        (rT := 3.4243, rA1 := 83.2821, rA2 := -78.0673, rA3 := 111.8853, rA4 := 0.3783, rA5 := 56.9060, rA6 := -96.9572),
        (rT := 3.5243, rA1 := 83.2822, rA2 := -77.8313, rA3 := 112.0983, rA4 := 0.2599, rA5 := 56.5349, rA6 := -96.8832),
        (rT := 3.6243, rA1 := 83.2821, rA2 := -77.6424, rA3 := 112.2616, rA4 := 0.2031, rA5 := 56.1792, rA6 := -96.8474),
        (rT := 3.7243, rA1 := 83.2821, rA2 := -77.4252, rA3 := 112.4477, rA4 := 0.1487, rA5 := 55.8068, rA6 := -96.8131),
        (rT := 3.8243, rA1 := 83.2821, rA2 := -77.2056, rA3 := 112.6319, rA4 := 0.1091, rA5 := 55.4161, rA6 := -96.7881),
        (rT := 3.9243, rA1 := 83.2821, rA2 := -76.9842, rA3 := 112.8135, rA4 := 0.0766, rA5 := 54.9796, rA6 := -96.7674),
        (rT := 4.0243, rA1 := 83.2821, rA2 := -76.7608, rA3 := 112.9927, rA4 := 0.0529, rA5 := 54.5444, rA6 := -96.7522),
        (rT := 4.1243, rA1 := 83.2821, rA2 := -76.4785, rA3 := 113.2129, rA4 := 0.0356, rA5 := 54.0667, rA6 := -96.7411),
        (rT := 4.2243, rA1 := 83.2821, rA2 := -76.3083, rA3 := 113.3440, rA4 := 0.0284, rA5 := 53.7920, rA6 := -96.7365),
        (* op 4 W10 - traj_robot2_W10 *)
        (rT := 0.0000, rA1 := 83.2821, rA2 := -76.3083, rA3 := 113.3440, rA4 := 0.0284, rA5 := 53.7920, rA6 := -96.7365),
        (rT := 0.2687, rA1 := 83.3426, rA2 := -76.2130, rA3 := 113.1677, rA4 := -0.8131, rA5 := 53.9876, rA6 := -96.2552),
        (rT := 0.5373, rA1 := 83.5109, rA2 := -75.9478, rA3 := 112.6767, rA4 := -3.1556, rA5 := 54.5321, rA6 := -94.9155),
        (rT := 0.8057, rA1 := 83.7674, rA2 := -75.5434, rA3 := 111.9284, rA4 := -6.7262, rA5 := 55.3620, rA6 := -92.8734),
        (rT := 1.0743, rA1 := 84.0926, rA2 := -75.0310, rA3 := 110.9799, rA4 := -11.2520, rA5 := 56.4139, rA6 := -90.2850),
        (rT := 1.3430, rA1 := 84.4668, rA2 := -74.4412, rA3 := 109.8884, rA4 := -16.4600, rA5 := 57.6244, rA6 := -87.3064),
        (rT := 1.6117, rA1 := 84.8705, rA2 := -73.8052, rA3 := 108.7111, rA4 := -22.0775, rA5 := 58.9300, rA6 := -84.0937),
        (rT := 1.8803, rA1 := 85.2839, rA2 := -73.1536, rA3 := 107.5052, rA4 := -27.8314, rA5 := 60.2673, rA6 := -80.8029),
        (rT := 2.1490, rA1 := 85.6875, rA2 := -72.5176, rA3 := 106.3279, rA4 := -33.4488, rA5 := 61.5730, rA6 := -77.5901),
        (rT := 2.4173, rA1 := 86.0617, rA2 := -71.9278, rA3 := 105.2364, rA4 := -38.6569, rA5 := 62.7835, rA6 := -74.6115),
        (rT := 2.6860, rA1 := 86.3869, rA2 := -71.4154, rA3 := 104.2879, rA4 := -43.1827, rA5 := 63.8354, rA6 := -72.0231),
        (rT := 2.9547, rA1 := 86.6434, rA2 := -71.0110, rA3 := 103.5396, rA4 := -46.7533, rA5 := 64.6653, rA6 := -69.9810),
        (rT := 3.2233, rA1 := 86.8118, rA2 := -70.7458, rA3 := 103.0487, rA4 := -49.0958, rA5 := 65.2097, rA6 := -68.6413),
        (rT := 3.4920, rA1 := 86.8722, rA2 := -70.6505, rA3 := 102.8723, rA4 := -49.9373, rA5 := 65.4053, rA6 := -68.1601),
        (rT := 3.5920, rA1 := 86.8724, rA2 := -70.2745, rA3 := 103.1990, rA4 := -50.2618, rA5 := 65.2813, rA6 := -67.7669),
        (rT := 3.6920, rA1 := 86.8725, rA2 := -69.7213, rA3 := 103.6748, rA4 := -50.7471, rA5 := 65.0552, rA6 := -67.1438),
        (rT := 3.7920, rA1 := 86.8726, rA2 := -69.4502, rA3 := 103.8964, rA4 := -51.0104, rA5 := 64.8316, rA6 := -66.7182),
        (rT := 3.8920, rA1 := 86.8725, rA2 := -69.2330, rA3 := 104.0648, rA4 := -51.2229, rA5 := 64.5888, rA6 := -66.3206),
        (rT := 3.9920, rA1 := 86.8725, rA2 := -68.9854, rA3 := 104.2549, rA4 := -51.4310, rA5 := 64.3399, rA6 := -65.9213),
        (rT := 4.0920, rA1 := 86.8725, rA2 := -68.7352, rA3 := 104.4418, rA4 := -51.6262, rA5 := 64.0843, rA6 := -65.5272),
        (rT := 4.1920, rA1 := 86.8725, rA2 := -68.4823, rA3 := 104.6258, rA4 := -51.8153, rA5 := 63.8254, rA6 := -65.1353),
        (rT := 4.2920, rA1 := 86.8725, rA2 := -68.2267, rA3 := 104.8067, rA4 := -51.9996, rA5 := 63.5638, rA6 := -64.7450),
        (rT := 4.3920, rA1 := 86.8725, rA2 := -67.9028, rA3 := 105.0279, rA4 := -52.2276, rA5 := 63.2357, rA6 := -64.2574),
        (rT := 4.4920, rA1 := 86.8725, rA2 := -67.7074, rA3 := 105.1595, rA4 := -52.3635, rA5 := 63.0382, rA6 := -63.9651),
        (* op 5 W11 - traj_robot2_W11 *)
        (rT := 0.0000, rA1 := 86.8725, rA2 := -67.7074, rA3 := 105.1595, rA4 := -52.3635, rA5 := 63.0382, rA6 := -63.9651),
        (rT := 0.2720, rA1 := 86.8241, rA2 := -67.7327, rA3 := 105.1314, rA4 := -51.4983, rA5 := 62.9127, rA6 := -64.4941),
        (rT := 0.5440, rA1 := 86.6893, rA2 := -67.8030, rA3 := 105.0531, rA4 := -49.0899, rA5 := 62.5634, rA6 := -65.9667),
        (rT := 0.8160, rA1 := 86.4839, rA2 := -67.9101, rA3 := 104.9338, rA4 := -45.4188, rA5 := 62.0309, rA6 := -68.2113),
        (rT := 1.0880, rA1 := 86.2236, rA2 := -68.0459, rA3 := 104.7826, rA4 := -40.7656, rA5 := 61.3560, rA6 := -71.0565),
        (rT := 1.3600, rA1 := 85.9240, rA2 := -68.2022, rA3 := 104.6086, rA4 := -35.4109, rA5 := 60.5793, rA6 := -74.3305),
        (rT := 1.6320, rA1 := 85.6008, rA2 := -68.3708, rA3 := 104.4209, rA4 := -29.6353, rA5 := 59.7416, rA6 := -77.8619),
        (rT := 1.9040, rA1 := 85.2698, rA2 := -68.5435, rA3 := 104.2287, rA4 := -23.7195, rA5 := 58.8836, rA6 := -81.4790),
        (rT := 2.1760, rA1 := 84.9467, rA2 := -68.7121, rA3 := 104.0410, rA4 := -17.9439, rA5 := 58.0459, rA6 := -85.0104),
        (rT := 2.4480, rA1 := 84.6471, rA2 := -68.8684, rA3 := 103.8670, rA4 := -12.5893, rA5 := 57.2692, rA6 := -88.2845),
        (rT := 2.7200, rA1 := 84.3867, rA2 := -69.0042, rA3 := 103.7158, rA4 := -7.9361, rA5 := 56.5943, rA6 := -91.1296),
        (rT := 2.9920, rA1 := 84.1813, rA2 := -69.1113, rA3 := 103.5965, rA4 := -4.2650, rA5 := 56.0618, rA6 := -93.3742),
        (rT := 3.2643, rA1 := 84.0465, rA2 := -69.1816, rA3 := 103.5183, rA4 := -1.8565, rA5 := 55.7125, rA6 := -94.8468),
        (rT := 3.5363, rA1 := 83.9981, rA2 := -69.2069, rA3 := 103.4901, rA4 := -0.9914, rA5 := 55.5870, rA6 := -95.3758),
        (rT := 3.6363, rA1 := 83.9979, rA2 := -68.8111, rA3 := 103.7925, rA4 := -0.7390, rA5 := 55.2565, rA6 := -95.5343),
        (rT := 3.7363, rA1 := 83.9975, rA2 := -68.2291, rA3 := 104.2324, rA4 := -0.3889, rA5 := 54.7233, rA6 := -95.7542),
        (rT := 3.8363, rA1 := 83.9975, rA2 := -67.9450, rA3 := 104.4363, rA4 := -0.2680, rA5 := 54.3464, rA6 := -95.8304),
        (rT := 3.9363, rA1 := 83.9975, rA2 := -67.7178, rA3 := 104.5907, rA4 := -0.2090, rA5 := 53.9648, rA6 := -95.8679),
        (rT := 4.0363, rA1 := 83.9975, rA2 := -67.4575, rA3 := 104.7656, rA4 := -0.1472, rA5 := 53.5219, rA6 := -95.9072),
        (rT := 4.1363, rA1 := 83.9975, rA2 := -67.1946, rA3 := 104.9375, rA4 := -0.1013, rA5 := 53.0634, rA6 := -95.9366),
        (rT := 4.2363, rA1 := 83.9976, rA2 := -66.9296, rA3 := 105.1060, rA4 := -0.0701, rA5 := 52.6202, rA6 := -95.9566),
        (rT := 4.3363, rA1 := 83.9976, rA2 := -66.6622, rA3 := 105.2713, rA4 := -0.0491, rA5 := 52.1805, rA6 := -95.9702),
        (rT := 4.4363, rA1 := 83.9976, rA2 := -66.3237, rA3 := 105.4730, rA4 := -0.0316, rA5 := 51.6342, rA6 := -95.9816),
        (rT := 4.5363, rA1 := 83.9976, rA2 := -66.1196, rA3 := 105.5927, rA4 := -0.0238, rA5 := 51.3075, rA6 := -95.9867),
        (* op 6 W12 - traj_robot2_W12 *)
        (rT := 0.0000, rA1 := 83.9976, rA2 := -66.1196, rA3 := 105.5927, rA4 := -0.0238, rA5 := 51.3075, rA6 := -95.9867),
        (rT := 0.2767, rA1 := 83.9002, rA2 := -66.1638, rA3 := 105.5263, rA4 := 0.8759, rA5 := 51.7354, rA6 := -96.4901),
        (rT := 0.5537, rA1 := 83.6309, rA2 := -66.2859, rA3 := 105.3425, rA4 := 3.3633, rA5 := 52.9183, rA6 := -97.8821),
        (rT := 0.8303, rA1 := 83.2241, rA2 := -66.4705, rA3 := 105.0648, rA4 := 7.1209, rA5 := 54.7054, rA6 := -99.9849),
        (rT := 1.1070, rA1 := 82.7141, rA2 := -66.7018, rA3 := 104.7167, rA4 := 11.8311, rA5 := 56.9455, rA6 := -102.6207),
        (rT := 1.3840, rA1 := 82.1354, rA2 := -66.9644, rA3 := 104.3218, rA4 := 17.1763, rA5 := 59.4877, rA6 := -105.6120),
        (rT := 1.6607, rA1 := 81.5224, rA2 := -67.2425, rA3 := 103.9033, rA4 := 22.8391, rA5 := 62.1808, rA6 := -108.7809),
        (rT := 1.9377, rA1 := 80.9093, rA2 := -67.5207, rA3 := 103.4849, rA4 := 28.5020, rA5 := 64.8740, rA6 := -111.9499),
        (rT := 2.2143, rA1 := 80.3306, rA2 := -67.7832, rA3 := 103.0899, rA4 := 33.8472, rA5 := 67.4162, rA6 := -114.9412),
        (rT := 2.4910, rA1 := 79.8207, rA2 := -68.0145, rA3 := 102.7418, rA4 := 38.5574, rA5 := 69.6563, rA6 := -117.5770),
        (rT := 2.7680, rA1 := 79.4138, rA2 := -68.1991, rA3 := 102.4642, rA4 := 42.3150, rA5 := 71.4433, rA6 := -119.6798),
        (rT := 3.0447, rA1 := 79.1446, rA2 := -68.3213, rA3 := 102.2804, rA4 := 44.8024, rA5 := 72.6263, rA6 := -121.0717),
        (rT := 3.3213, rA1 := 79.0472, rA2 := -68.3655, rA3 := 102.2139, rA4 := 45.7021, rA5 := 73.0542, rA6 := -121.5752),
        (rT := 3.4213, rA1 := 79.0469, rA2 := -67.9761, rA3 := 102.5143, rA4 := 45.9316, rA5 := 72.9480, rA6 := -121.8853),
        (rT := 3.5213, rA1 := 79.0466, rA2 := -67.4036, rA3 := 102.9515, rA4 := 46.2710, rA5 := 72.7498, rA6 := -122.3762),
        (rT := 3.6213, rA1 := 79.0465, rA2 := -67.1241, rA3 := 103.1540, rA4 := 46.4436, rA5 := 72.5500, rA6 := -122.7036),
        (rT := 3.7213, rA1 := 79.0466, rA2 := -66.9006, rA3 := 103.3074, rA4 := 46.5817, rA5 := 72.3183, rA6 := -123.0218),
        (rT := 3.8213, rA1 := 79.0466, rA2 := -66.6446, rA3 := 103.4812, rA4 := 46.7318, rA5 := 72.0473, rA6 := -123.3823),
        (rT := 3.9213, rA1 := 79.0466, rA2 := -66.3860, rA3 := 103.6520, rA4 := 46.8746, rA5 := 71.7590, rA6 := -123.7488),
        (rT := 4.0213, rA1 := 79.0466, rA2 := -66.1253, rA3 := 103.8194, rA4 := 47.0062, rA5 := 71.4712, rA6 := -124.1033),
        (rT := 4.1213, rA1 := 79.0466, rA2 := -65.8625, rA3 := 103.9835, rA4 := 47.1279, rA5 := 71.1891, rA6 := -124.4433),
        (rT := 4.2213, rA1 := 79.0466, rA2 := -65.5304, rA3 := 104.1833, rA4 := 47.2638, rA5 := 70.8638, rA6 := -124.8302),
        (rT := 4.3213, rA1 := 79.0466, rA2 := -65.3303, rA3 := 104.3019, rA4 := 47.3413, rA5 := 70.6741, rA6 := -125.0540),
        (* op 7 W09 - traj_robot2_W09 *)
        (rT := 0.0000, rA1 := 79.0466, rA2 := -65.3303, rA3 := 104.3019, rA4 := 47.3413, rA5 := 70.6741, rA6 := -125.0540),
        (rT := 0.2997, rA1 := 79.2593, rA2 := -64.3494, rA3 := 101.6347, rA4 := 47.1082, rA5 := 71.5396, rA6 := -123.8549),
        (rT := 0.5993, rA1 := 79.7271, rA2 := -62.1915, rA3 := 95.7668, rA4 := 46.5953, rA5 := 73.4437, rA6 := -121.2168),
        (rT := 0.8990, rA1 := 80.1949, rA2 := -60.0336, rA3 := 89.8989, rA4 := 46.0825, rA5 := 75.3478, rA6 := -118.5786),
        (rT := 1.1987, rA1 := 80.4076, rA2 := -59.0528, rA3 := 87.2316, rA4 := 45.8493, rA5 := 76.2133, rA6 := -117.3795),
        (rT := 1.2987, rA1 := 80.4077, rA2 := -58.7325, rA3 := 87.5160, rA4 := 45.8400, rA5 := 76.2458, rA6 := -117.3487),
        (rT := 1.3987, rA1 := 80.4079, rA2 := -58.2594, rA3 := 87.9317, rA4 := 45.8493, rA5 := 76.2133, rA6 := -117.3795),
        (rT := 1.4987, rA1 := 80.4079, rA2 := -58.0224, rA3 := 88.1304, rA4 := 45.9151, rA5 := 75.9863, rA6 := -117.5926),
        (rT := 1.5987, rA1 := 80.4079, rA2 := -57.8310, rA3 := 88.2828, rA4 := 45.9995, rA5 := 75.6941, rA6 := -117.8717),
        (rT := 1.6987, rA1 := 80.4079, rA2 := -57.6175, rA3 := 88.4503, rA4 := 46.0740, rA5 := 75.4333, rA6 := -118.1321),
        (rT := 1.7987, rA1 := 80.4079, rA2 := -57.4030, rA3 := 88.6137, rA4 := 46.1486, rA5 := 75.1723, rA6 := -118.3992),
        (rT := 1.8987, rA1 := 80.4079, rA2 := -57.1859, rA3 := 88.7745, rA4 := 46.2237, rA5 := 74.9116, rA6 := -118.6705),
        (rT := 1.9987, rA1 := 80.4079, rA2 := -56.9666, rA3 := 88.9322, rA4 := 46.2996, rA5 := 74.6512, rA6 := -118.9454),
        (rT := 2.0987, rA1 := 80.4079, rA2 := -56.6891, rA3 := 89.1244, rA4 := 46.3958, rA5 := 74.3266, rA6 := -119.2925),
        (rT := 2.1987, rA1 := 80.4079, rA2 := -56.5217, rA3 := 89.2385, rA4 := 46.4540, rA5 := 74.1321, rA6 := -119.5017),
        (* op 8 W08 - traj_robot2_W08 *)
        (rT := 0.0000, rA1 := 80.4079, rA2 := -56.5217, rA3 := 89.2385, rA4 := 46.4540, rA5 := 74.1321, rA6 := -119.5017),
        (rT := 0.2813, rA1 := 80.5091, rA2 := -56.5983, rA3 := 89.2213, rA4 := 45.3937, rA5 := 73.8342, rA6 := -118.9496),
        (rT := 0.5627, rA1 := 80.7866, rA2 := -56.8083, rA3 := 89.1743, rA4 := 42.4866, rA5 := 73.0173, rA6 := -117.4358),
        (rT := 0.8437, rA1 := 81.2013, rA2 := -57.1220, rA3 := 89.1041, rA4 := 38.1430, rA5 := 71.7968, rA6 := -115.1739),
        (rT := 1.1250, rA1 := 81.7139, rA2 := -57.5099, rA3 := 89.0173, rA4 := 32.7734, rA5 := 70.2880, rA6 := -112.3778),
        (rT := 1.4063, rA1 := 82.2852, rA2 := -57.9422, rA3 := 88.9205, rA4 := 26.7881, rA5 := 68.6061, rA6 := -109.2610),
        (rT := 1.6877, rA1 := 82.8762, rA2 := -58.3894, rA3 := 88.8205, rA4 := 20.5976, rA5 := 66.8666, rA6 := -106.0374),
        (rT := 1.9687, rA1 := 83.4476, rA2 := -58.8217, rA3 := 88.7237, rA4 := 14.6124, rA5 := 65.1848, rA6 := -102.9207),
        (rT := 2.2500, rA1 := 83.9602, rA2 := -59.2095, rA3 := 88.6369, rA4 := 9.2428, rA5 := 63.6760, rA6 := -100.1245),
        (rT := 2.5313, rA1 := 84.3749, rA2 := -59.5233, rA3 := 88.5667, rA4 := 4.8992, rA5 := 62.4554, rA6 := -97.8626),
        (rT := 2.8127, rA1 := 84.6524, rA2 := -59.7333, rA3 := 88.5197, rA4 := 1.9920, rA5 := 61.6386, rA6 := -96.3488),
        (rT := 3.0940, rA1 := 84.7536, rA2 := -59.8099, rA3 := 88.5026, rA4 := 0.9318, rA5 := 61.3406, rA6 := -95.7967),
        (rT := 3.1940, rA1 := 84.7538, rA2 := -59.4813, rA3 := 88.7926, rA4 := 0.7130, rA5 := 61.0466, rA6 := -95.6684),
        (rT := 3.2940, rA1 := 84.7541, rA2 := -58.9980, rA3 := 89.2147, rA4 := 0.4049, rA5 := 60.5635, rA6 := -95.4875),
        (rT := 3.3940, rA1 := 84.7542, rA2 := -58.7611, rA3 := 89.4106, rA4 := 0.2844, rA5 := 60.1937, rA6 := -95.4165),
        (rT := 3.4940, rA1 := 84.7541, rA2 := -58.5715, rA3 := 89.5589, rA4 := 0.2172, rA5 := 59.8274, rA6 := -95.3767),
        (rT := 3.5940, rA1 := 84.7541, rA2 := -58.3554, rA3 := 89.7259, rA4 := 0.1585, rA5 := 59.4538, rA6 := -95.3418),
        (rT := 3.6940, rA1 := 84.7541, rA2 := -58.1373, rA3 := 89.8898, rA4 := 0.1165, rA5 := 59.0779, rA6 := -95.3167),
        (rT := 3.7940, rA1 := 84.7541, rA2 := -57.9170, rA3 := 90.0506, rA4 := 0.0850, rA5 := 58.7008, rA6 := -95.2978),
        (rT := 3.8940, rA1 := 84.7541, rA2 := -57.6945, rA3 := 90.2085, rA4 := 0.0625, rA5 := 58.3229, rA6 := -95.2842),
        (rT := 3.9940, rA1 := 84.7541, rA2 := -57.4129, rA3 := 90.4008, rA4 := 0.0429, rA5 := 57.8503, rA6 := -95.2723),
        (rT := 4.0940, rA1 := 84.7541, rA2 := -57.2430, rA3 := 90.5150, rA4 := 0.0336, rA5 := 57.5666, rA6 := -95.2667),
        (* op 9 W07 - traj_robot2_W07 *)
        (rT := 0.0000, rA1 := 84.7541, rA2 := -57.2430, rA3 := 90.5150, rA4 := 0.0336, rA5 := 57.5666, rA6 := -95.2667),
        (rT := 0.2723, rA1 := 84.8408, rA2 := -57.2997, rA3 := 90.4856, rA4 := -0.9166, rA5 := 57.7929, rA6 := -94.7597),
        (rT := 0.5450, rA1 := 85.0806, rA2 := -57.4562, rA3 := 90.4044, rA4 := -3.5434, rA5 := 58.4188, rA6 := -93.3581),
        (rT := 0.8173, rA1 := 85.4427, rA2 := -57.6927, rA3 := 90.2817, rA4 := -7.5116, rA5 := 59.3642, rA6 := -91.2408),
        (rT := 1.0897, rA1 := 85.8967, rA2 := -57.9891, rA3 := 90.1280, rA4 := -12.4859, rA5 := 60.5494, rA6 := -88.5867),
        (rT := 1.3623, rA1 := 86.4118, rA2 := -58.3255, rA3 := 89.9535, rA4 := -18.1308, rA5 := 61.8943, rA6 := -85.5747),
        (rT := 1.6347, rA1 := 86.9576, rA2 := -58.6819, rA3 := 89.7687, rA4 := -24.1111, rA5 := 63.3191, rA6 := -82.3838),
        (rT := 1.9070, rA1 := 87.5034, rA2 := -59.0383, rA3 := 89.5838, rA4 := -30.0914, rA5 := 64.7440, rA6 := -79.1929),
        (rT := 2.1797, rA1 := 88.0186, rA2 := -59.3747, rA3 := 89.4093, rA4 := -35.7363, rA5 := 66.0889, rA6 := -76.1810),
        (rT := 2.4520, rA1 := 88.4725, rA2 := -59.6712, rA3 := 89.2556, rA4 := -40.7106, rA5 := 67.2740, rA6 := -73.5268),
        (rT := 2.7243, rA1 := 88.8347, rA2 := -59.9076, rA3 := 89.1329, rA4 := -44.6788, rA5 := 68.2195, rA6 := -71.4095),
        (rT := 2.9970, rA1 := 89.0744, rA2 := -60.0642, rA3 := 89.0517, rA4 := -47.3057, rA5 := 68.8453, rA6 := -70.0079),
        (rT := 3.2693, rA1 := 89.1611, rA2 := -60.1208, rA3 := 89.0224, rA4 := -48.2558, rA5 := 69.0717, rA6 := -69.5010),
        (rT := 3.3693, rA1 := 89.1614, rA2 := -59.7902, rA3 := 89.3125, rA4 := -48.5199, rA5 := 68.9754, rA6 := -69.1961),
        (rT := 3.4693, rA1 := 89.1617, rA2 := -59.3039, rA3 := 89.7347, rA4 := -48.9126, rA5 := 68.7948, rA6 := -68.7101),
        (rT := 3.5693, rA1 := 89.1617, rA2 := -59.0656, rA3 := 89.9307, rA4 := -49.1199, rA5 := 68.6061, rA6 := -68.3719),
        (rT := 3.6693, rA1 := 89.1616, rA2 := -58.8747, rA3 := 90.0789, rA4 := -49.2838, rA5 := 68.3967, rA6 := -68.0517),
        (rT := 3.7693, rA1 := 89.1616, rA2 := -58.6574, rA3 := 90.2460, rA4 := -49.4444, rA5 := 68.1793, rA6 := -67.7272),
        (rT := 3.8693, rA1 := 89.1616, rA2 := -58.4380, rA3 := 90.4100, rA4 := -49.5935, rA5 := 67.9536, rA6 := -67.4047),
        (rT := 3.9693, rA1 := 89.1616, rA2 := -58.2163, rA3 := 90.5709, rA4 := -49.7362, rA5 := 67.7230, rA6 := -67.0834),
        (rT := 4.0693, rA1 := 89.1616, rA2 := -57.9925, rA3 := 90.7288, rA4 := -49.8734, rA5 := 67.4885, rA6 := -66.7630),
        (rT := 4.1693, rA1 := 89.1616, rA2 := -57.7091, rA3 := 90.9212, rA4 := -50.0409, rA5 := 67.1925, rA6 := -66.3631),
        (rT := 4.2693, rA1 := 89.1616, rA2 := -57.5383, rA3 := 91.0354, rA4 := -50.1401, rA5 := 67.0139, rA6 := -66.1234),
        (* op 10 HOME - traj_robot2_n26 *)
        (rT := 0.0000, rA1 := 89.1616, rA2 := -57.5383, rA3 := 91.0354, rA4 := -50.1401, rA5 := 67.0139, rA6 := -66.1234),
        (rT := 0.2010, rA1 := 88.8893, rA2 := -57.6374, rA3 := 91.0323, rA4 := -49.9869, rA5 := 66.8092, rA6 := -65.9214),
        (rT := 0.4020, rA1 := 88.0961, rA2 := -57.9262, rA3 := 91.0231, rA4 := -49.5409, rA5 := 66.2131, rA6 := -65.3332),
        (rT := 0.6028, rA1 := 86.8182, rA2 := -58.3915, rA3 := 91.0082, rA4 := -48.8222, rA5 := 65.2526, rA6 := -64.3854),
        (rT := 0.8037, rA1 := 85.0913, rA2 := -59.0202, rA3 := 90.9882, rA4 := -47.8511, rA5 := 63.9546, rA6 := -63.1048),
        (rT := 1.0047, rA1 := 82.9513, rA2 := -59.7993, rA3 := 90.9633, rA4 := -46.6477, rA5 := 62.3463, rA6 := -61.5178),
        (rT := 1.2057, rA1 := 80.4343, rA2 := -60.7157, rA3 := 90.9341, rA4 := -45.2323, rA5 := 60.4545, rA6 := -59.6511),
        (rT := 1.4065, rA1 := 77.5761, rA2 := -61.7563, rA3 := 90.9009, rA4 := -43.6249, rA5 := 58.3062, rA6 := -57.5314),
        (rT := 1.6075, rA1 := 74.4126, rA2 := -62.9081, rA3 := 90.8642, rA4 := -41.8459, rA5 := 55.9285, rA6 := -55.1853),
        (rT := 1.8085, rA1 := 70.9797, rA2 := -64.1579, rA3 := 90.8243, rA4 := -39.9155, rA5 := 53.3484, rA6 := -52.6395),
        (rT := 2.0095, rA1 := 67.3134, rA2 := -65.4927, rA3 := 90.7817, rA4 := -37.8537, rA5 := 50.5928, rA6 := -49.9205),
        (rT := 2.2105, rA1 := 63.4496, rA2 := -66.8995, rA3 := 90.7368, rA4 := -35.6809, rA5 := 47.6887, rA6 := -47.0550),
        (rT := 2.4112, rA1 := 59.4241, rA2 := -68.3650, rA3 := 90.6901, rA4 := -33.4172, rA5 := 44.6632, rA6 := -44.0697),
        (rT := 2.6122, rA1 := 55.2730, rA2 := -69.8764, rA3 := 90.6419, rA4 := -31.0828, rA5 := 41.5432, rA6 := -40.9911),
        (rT := 2.8132, rA1 := 51.0320, rA2 := -71.4204, rA3 := 90.5926, rA4 := -28.6979, rA5 := 38.3557, rA6 := -37.8460),
        (rT := 3.0142, rA1 := 46.7372, rA2 := -72.9841, rA3 := 90.5428, rA4 := -26.2827, rA5 := 35.1277, rA6 := -34.6609),
        (rT := 3.2150, rA1 := 42.4244, rA2 := -74.5542, rA3 := 90.4927, rA4 := -23.8574, rA5 := 31.8862, rA6 := -31.4625),
        (rT := 3.4160, rA1 := 38.1296, rA2 := -76.1179, rA3 := 90.4428, rA4 := -21.4422, rA5 := 28.6582, rA6 := -28.2774),
        (rT := 3.6170, rA1 := 33.8887, rA2 := -77.6619, rA3 := 90.3935, rA4 := -19.0573, rA5 := 25.4707, rA6 := -25.1323),
        (rT := 3.8180, rA1 := 29.7375, rA2 := -79.1733, rA3 := 90.3453, rA4 := -16.7229, rA5 := 22.3507, rA6 := -22.0537),
        (rT := 4.0190, rA1 := 25.7120, rA2 := -80.6388, rA3 := 90.2986, rA4 := -14.4592, rA5 := 19.3252, rA6 := -19.0684),
        (rT := 4.2197, rA1 := 21.8482, rA2 := -82.0456, rA3 := 90.2537, rA4 := -12.2863, rA5 := 16.4211, rA6 := -16.2029),
        (rT := 4.4207, rA1 := 18.1819, rA2 := -83.3804, rA3 := 90.2111, rA4 := -10.2246, rA5 := 13.6655, rA6 := -13.4839),
        (rT := 4.6217, rA1 := 14.7490, rA2 := -84.6302, rA3 := 90.1713, rA4 := -8.2941, rA5 := 11.0854, rA6 := -10.9381),
        (rT := 4.8228, rA1 := 11.5855, rA2 := -85.7820, rA3 := 90.1345, rA4 := -6.5151, rA5 := 8.7077, rA6 := -8.5920),
        (rT := 5.0235, rA1 := 8.7273, rA2 := -86.8226, rA3 := 90.1014, rA4 := -4.9078, rA5 := 6.5594, rA6 := -6.4723),
        (rT := 5.2245, rA1 := 6.2103, rA2 := -87.7390, rA3 := 90.0721, rA4 := -3.4924, rA5 := 4.6676, rA6 := -4.6056),
        (rT := 5.4255, rA1 := 4.0704, rA2 := -88.5181, rA3 := 90.0473, rA4 := -2.2890, rA5 := 3.0593, rA6 := -3.0186),
        (rT := 5.6265, rA1 := 2.3434, rA2 := -89.1468, rA3 := 90.0272, rA4 := -1.3178, rA5 := 1.7613, rA6 := -1.7379),
        (rT := 5.8275, rA1 := 1.0655, rA2 := -89.6121, rA3 := 90.0124, rA4 := -0.5992, rA5 := 0.8008, rA6 := -0.7902),
        (rT := 6.0282, rA1 := 0.2724, rA2 := -89.9008, rA3 := 90.0032, rA4 := -0.1532, rA5 := 0.2047, rA6 := -0.2020),
        (rT := 6.2292, rA1 := 0.0000, rA2 := -90.0000, rA3 := 90.0000, rA4 := 0.0000, rA5 := 0.0000, rA6 := 0.0000)
    ];
END_VAR
END_NAMESPACE

(* ---- FB_JointAngleEncoder.st ---- *)
(*
 * FB_JointAngleEncoder
 * Device simulator R2 (robot2), cell welding_cell_2_small. Generated by bt2plc 0.1.0.
 *
 * Encodes six KUKA robot joint angles (REAL degrees) into the VASS Option area
 * as scaled fixed-point INTs (0.02 deg per count, big-endian byte order).
 *
 * Encoding per encoding.md:
 *   count = ROUND(angle_deg / 0.02)   clamped to [-32768, +32767]
 *   Byte layout: big-endian (high byte first) in each 2-byte pair
 *
 * Output abyOption = Option area aVassInputData[16..27], 2 bytes per axis
 * (PLC_PRG copies it into the robot -> PLC telegram):
 *   abyOption[0-1]  = bytes 16-17 = A1,  abyOption[2-3]   = bytes 18-19 = A2,
 *   abyOption[4-5]  = bytes 20-21 = A3,  abyOption[6-7]   = bytes 22-23 = A4,
 *   abyOption[8-9]  = bytes 24-25 = A5,  abyOption[10-11] = bytes 26-27 = A6
 *)

FUNCTION_BLOCK FB_JointAngleEncoder
VAR_INPUT
    rA1_deg     : REAL := 0.0;      (* Axis 1 angle in degrees *)
    rA2_deg     : REAL := 0.0;      (* Axis 2 angle in degrees *)
    rA3_deg     : REAL := 0.0;      (* Axis 3 angle in degrees *)
    rA4_deg     : REAL := 0.0;      (* Axis 4 angle in degrees *)
    rA5_deg     : REAL := 0.0;      (* Axis 5 angle in degrees *)
    rA6_deg     : REAL := 0.0;      (* Axis 6 angle in degrees *)
END_VAR

VAR_OUTPUT
    (* Encoded INT values (for monitoring/debug) *)
    iA1_count   : INT;
    iA2_count   : INT;
    iA3_count   : INT;
    iA4_count   : INT;
    iA5_count   : INT;
    iA6_count   : INT;

    (* Option area bytes 16..27 of the robot -> PLC telegram, big-endian A1..A6 *)
    abyOption   : ARRAY[0..11] OF BYTE;
END_VAR

VAR CONSTANT
    SCALE_FACTOR    : REAL := 0.02;     (* degrees per count *)
    INV_SCALE       : REAL := 50.0;     (* 1/0.02 = 50, multiply for speed *)
    COUNT_MAX       : DINT := 32767;
    COUNT_MIN       : DINT := -32768;
END_VAR

VAR
    _arDeg      : ARRAY[1..6] OF REAL;
    _aiCount    : ARRAY[1..6] OF INT;
    _diTemp     : DINT;
    _wTemp      : WORD;
    _i          : INT;
END_VAR
(*
 * FB_JointAngleEncoder - Implementation
 *
 * Converts 6x REAL degree angles to scaled INT counts (0.02 deg per count)
 * and writes them big-endian into abyOption[0..11] (telegram bytes 16..27).
 *
 * Conversion:  count = ROUND(angle / 0.02)  clamped to INT range
 * Byte order:  Big-endian (high byte at lower address) per S7/PROFINET convention
 * Two's complement is formed in DINT (count + 65536 for negative counts), so no
 * bit operation is applied to a signed type.
 *)

_arDeg[1] := rA1_deg;
_arDeg[2] := rA2_deg;
_arDeg[3] := rA3_deg;
_arDeg[4] := rA4_deg;
_arDeg[5] := rA5_deg;
_arDeg[6] := rA6_deg;

FOR _i := 1 TO 6 DO
    (* === Scale and clamp === *)
    _diTemp := REAL_TO_DINT(LIMIT(REAL#-32768.0, _arDeg[_i] * INV_SCALE, REAL#32767.0));
    IF _diTemp > COUNT_MAX THEN _diTemp := COUNT_MAX; END_IF
    IF _diTemp < COUNT_MIN THEN _diTemp := COUNT_MIN; END_IF
    _aiCount[_i] := DINT_TO_INT(_diTemp);

    (* === Big-endian into the Option area: high byte first === *)
    IF _diTemp < 0 THEN
        _diTemp := _diTemp + 65536;
    END_IF
    _wTemp := DINT_TO_WORD(_diTemp);
    abyOption[2 * (_i - 1)] := WORD_TO_BYTE(SHR(_wTemp, 8));
    abyOption[2 * (_i - 1) + 1] := WORD_TO_BYTE(_wTemp AND WORD#16#FF);
END_FOR

iA1_count := _aiCount[1];
iA2_count := _aiCount[2];
iA3_count := _aiCount[3];
iA4_count := _aiCount[4];
iA5_count := _aiCount[5];
iA6_count := _aiCount[6];
END_FUNCTION_BLOCK

(* ---- FB_PROFIsafe_Simulator.st ---- *)
(*
 * FB_PROFIsafe_Simulator
 * Device simulator R2 (robot2), cell welding_cell_2_small. Generated by bt2plc 0.1.0.
 *
 * Simulates the PROFIsafe protocol layer for the FDIO64 module (Slot 1).
 * In a real KUKA controller, the PROFIsafe stack handles CRC generation,
 * sequence counters, and watchdog monitoring.
 *
 * For simulation purposes, this FB:
 * - Monitors the safe output bytes from the PLC (abySafeOut = copy of GVL_IO.bySafeOut0..7)
 * - Provides a "communication OK" flag
 *
 * IMPORTANT: This does NOT provide real functional safety!
 * It only generates data patterns that allow the PLC's PROFIsafe stack
 * to accept the device as communicating. For real safety testing,
 * you need a certified PROFIsafe device or test equipment.
 *
 * PROFIsafe frame structure per IEC 61784-3-3:
 *   [User Data (8 bytes)] [Status/Control (1 byte)] [CRC (3 bytes)]
 *
 * Status byte bits (F_Input from device):
 *   Bit 0: Toggle bit (alternates each cycle)
 *   Bit 1: Reserved
 *   Bit 2: Data valid
 *   Bit 3-7: Reserved / Sequence counter
 *
 * Control byte bits (F_Output from controller):
 *   Bit 0: Toggle bit
 *   Bit 1: Activate device
 *   Bit 2: Reserved
 *   Bit 3-7: Reserved
 *)

FUNCTION_BLOCK FB_PROFIsafe_Simulator
VAR_INPUT
    bEnable         : BOOL := TRUE;
    dwF_Source_Add  : DWORD := DWORD#1;     (* F_Source_Add from parameterization *)
    dwF_Dest_Add    : DWORD := DWORD#1;     (* F_Dest_Add from parameterization *)
    tF_WD_Time      : TIME := T#500MS;      (* Watchdog time *)
    abySafeOut      : ARRAY[0..7] OF BYTE;  (* Safe outputs PLC -> robot (GVL_IO.bySafeOut0..7) *)
END_VAR

VAR_OUTPUT
    bCommOK         : BOOL;                 (* PROFIsafe communication established *)
    bDataValid      : BOOL;                 (* Safe data is valid *)
    bWatchdogError  : BOOL;                 (* Watchdog timeout *)
END_VAR

VAR
    _bToggleBit     : BOOL;                 (* Toggle bit for sequence *)
    _nSeqCounter    : BYTE;                 (* Sequence counter 0-31 *)
    _nCycleCount    : UDINT;                (* Absolute cycle counter *)

    (* Watchdog *)
    _tonWatchdog    : TON;
    _bPLCSafeActive : BOOL;

    (* CRC calculation helper *)
    _dwCrcSeed      : DWORD;
END_VAR
(*
 * FB_PROFIsafe_Simulator - Implementation
 * Works on the input image abySafeOut (PLC_PRG copies GVL_IO.bySafeOut0..7).
 *)

IF NOT bEnable THEN
    bCommOK := FALSE;
    bDataValid := FALSE;
    RETURN;
END_IF

IF _nCycleCount < UDINT#4000000000 THEN
    _nCycleCount := _nCycleCount + 1;
ELSE
    _nCycleCount := 0;
END_IF

(* ============================================================================
   MONITOR PLC SAFE OUTPUT DATA
   ============================================================================ *)
_bPLCSafeActive := (abySafeOut[0] <> BYTE#0) OR (abySafeOut[1] <> BYTE#0);

(* Watchdog *)
_tonWatchdog(IN := NOT _bPLCSafeActive, PT := tF_WD_Time);
bWatchdogError := _tonWatchdog.Q;

bCommOK := _bPLCSafeActive AND NOT bWatchdogError;
bDataValid := bCommOK;
END_FUNCTION_BLOCK

(* ---- FB_ProgramPlayer.st ---- *)
(*
 * FB_ProgramPlayer
 * Device simulator R2 (robot2), cell welding_cell_2_small, tree bt_1790934549_welding_cell_2_small. Generated by bt2plc 0.1.0.
 *
 * Plays the bt2plc robot program (GVL_Program) for PROD_FOLGE, or a blind joint
 * move to the home pose for HOME_FOLGE. Robot side of the zone protocol, per op k
 * with mask M = GVL_Program.aOps[k].dwZoneMask:
 *   1  wStep := k                          (also for M = 0)
 *   2  if M <> 0: REQUEST := M             (same call / telegram as wStep)
 *   3  if M <> 0: wait (GRANT AND M) = M
 *   4  start delay; trajectory (x rVelScale x override); hold
 *   5  if M <> 0: REQUEST := 0
 *   6  if M <> 0: wait (GRANT AND M) = 0   (4-phase, before the next REQUEST)
 *   7  next op; after the last op: bDone, wStep := 0 (same call)
 *
 * Timing: all times are REAL seconds accumulated from rDt (seconds per call, the
 * device task interval). Motion time advances by rDt * rRate * rVelScale, delay and
 * hold by rDt (the override does not scale dwell times). No TIME() / TON is used.
 * Zero-time transitions fall through within one call (at most N_MAX_TRANSITIONS),
 * but wStep changes at most once per call, so every step is visible to the head PLC.
 * Joints (deg) are linearly interpolated between waypoints and published as rA1..rA6_deg.
 * Abort (bAbort level while busy): REQUEST := 0, wStep := 0, the pose is held.
 * The robot powers up at GVL_Program.arHomeDeg.
 *)

FUNCTION_BLOCK FB_ProgramPlayer
VAR_INPUT
    bStart          : BOOL;                 (* Rising edge: start wJob *)
    wJob            : WORD;                 (* Folge to play: PROD_FOLGE or HOME_FOLGE *)
    bAbort          : BOOL;                 (* Level: stop / cancel / drives off / E-stop *)
    dwGrant         : DWORD;                (* Zone GRANT bits from the head PLC *)
    rRate           : REAL := 1.0;          (* Speed override factor (1.0 = 100 %) *)
    rDt             : REAL := 0.02;         (* Seconds per call (task interval) *)
END_VAR

VAR_OUTPUT
    eState          : E_PlayerState;        (* Current state *)
    bBusy           : BOOL;                 (* Program running *)
    bDone           : BOOL;                 (* Latched until next start *)
    bError          : BOOL;                 (* Latched until next start *)
    wErrorCode      : WORD;                 (* Error code, GVL_Program.ERR_xxx *)
    wWarningCode    : WORD;                 (* Warning code, GVL_Program.WARN_xxx, latched until next start *)
    wStep           : WORD;                 (* 1-based op index, 0 = none *)
    dwRequest       : DWORD;                (* Zone REQUEST bits to the head PLC *)
    bAtHome         : BOOL;                 (* All joints within R_AT_HOME_TOL_DEG of arHomeDeg *)
    rA1_deg         : REAL;                 (* Axis 1 angle *)
    rA2_deg         : REAL;                 (* Axis 2 angle *)
    rA3_deg         : REAL;                 (* Axis 3 angle *)
    rA4_deg         : REAL;                 (* Axis 4 angle *)
    rA5_deg         : REAL;                 (* Axis 5 angle *)
    rA6_deg         : REAL;                 (* Axis 6 angle *)
END_VAR

VAR CONSTANT
    N_MAX_TRANSITIONS : INT := 8;           (* Fall-through bound per call *)
END_VAR

VAR
    _eState         : E_PlayerState := E_PlayerState#PS_IDLE;
    _rtrigStart     : R_TRIG;
    _bFirstCall     : BOOL := TRUE;

    (* === Current op === *)
    _nOp            : INT;                  (* 1-based op index, 0 = HOME_FOLGE move *)
    _dwMask         : DWORD;                (* Zone mask of the current op *)
    _bHomeMove      : BOOL;                 (* Current move is a blind home move *)
    _nWp            : INT;                  (* Current waypoint segment start *)
    _nLast          : INT;                  (* Last waypoint of the current op, 0 = none *)
    _rVel           : REAL;                 (* Velocity scale of the current move *)

    (* === Time (s) === *)
    _rDtCall        : REAL;                 (* rDt limited to 0..1 s *)
    _rRateCall      : REAL;                 (* rRate limited to >= 0 *)
    _rT             : REAL;                 (* Motion time since move start *)
    _rTimer         : REAL;                 (* Delay / hold timer *)
    _rDur           : REAL;                 (* Duration of the blind home move *)
    _rAlpha         : REAL;                 (* Interpolation factor 0..1 *)
    _rSpan          : REAL;                 (* Waypoint segment duration *)

    (* === Pose (deg) === *)
    _arQ            : ARRAY[1..6] OF REAL;  (* Current joint angles *)
    _arQ0           : ARRAY[1..6] OF REAL;  (* Pose at the start of a blind home move *)
    _arQa           : ARRAY[1..6] OF REAL;  (* Segment start waypoint *)
    _arQb           : ARRAY[1..6] OF REAL;  (* Segment end waypoint *)

    (* === Fall-through === *)
    _nPass          : INT;
    _bAdvance       : BOOL;                 (* A transition happened in this pass *)
    _bStepSet       : BOOL;                 (* wStep changed in this call *)
    _bMoveDone      : BOOL;
    _i              : INT;
END_VAR
(*
 * FB_ProgramPlayer - Implementation
 *)

(* ============================================================================
   INIT - the robot powers up at the home pose
   ============================================================================ *)
IF _bFirstCall THEN
    FOR _i := 1 TO 6 DO
        _arQ[_i] := GVL_Program.arHomeDeg[_i];
    END_FOR
    _bFirstCall := FALSE;
END_IF

_rDtCall := LIMIT(0.0, rDt, 1.0);
_rRateCall := MAX(rRate, 0.0);
_rtrigStart(CLK := bStart);

(* ============================================================================
   ABORT - stop / cancel / drives off / E-stop: REQUEST := 0, wStep := 0, hold pose
   ============================================================================ *)
IF bAbort AND bBusy THEN
    _eState := E_PlayerState#PS_IDLE;
    bBusy := FALSE;
    wStep := WORD#0;
    dwRequest := DWORD#0;
END_IF

(* ============================================================================
   CLOCK - advance the timer of the state that is active at the start of the call
   (a state entered during this call starts counting with the next call)
   ============================================================================ *)
IF _eState = E_PlayerState#PS_DELAY OR _eState = E_PlayerState#PS_HOLD THEN
    _rTimer := _rTimer + _rDtCall;
ELSIF _eState = E_PlayerState#PS_MOVE THEN
    _rT := _rT + _rDtCall * _rRateCall * _rVel;
END_IF

(* ============================================================================
   START
   ============================================================================ *)
IF _rtrigStart.Q AND NOT bBusy AND NOT bAbort THEN
    bDone := FALSE;
    bError := FALSE;
    wErrorCode := WORD#0;
    wWarningCode := WORD#0;
    wStep := WORD#0;
    dwRequest := DWORD#0;
    _nOp := 0;
    _dwMask := DWORD#0;
    _rT := 0.0;
    _rTimer := 0.0;
    IF wJob = GVL_Program.HOME_FOLGE THEN
        (* Blind joint move from the current pose to arHomeDeg: no step, no zones *)
        FOR _i := 1 TO 6 DO
            _arQ0[_i] := _arQ[_i];
        END_FOR
        _bHomeMove := TRUE;
        _nLast := 0;
        _rVel := 1.0;
        _rDur := GVL_Program.R_HOME_S;
        bBusy := TRUE;
        _eState := E_PlayerState#PS_MOVE;
    ELSIF wJob = GVL_Program.PROD_FOLGE AND GVL_Program.N_OPS > 0 THEN
        bBusy := TRUE;
        _eState := E_PlayerState#PS_NEXT_OP;
    ELSE
        wErrorCode := GVL_Program.ERR_UNKNOWN_FOLGE;
        _eState := E_PlayerState#PS_ERROR;
    END_IF
END_IF

(* ============================================================================
   STATE MACHINE - falls through zero-time transitions (bounded)
   ============================================================================ *)
_bStepSet := FALSE;
FOR _nPass := 1 TO N_MAX_TRANSITIONS DO
    _bAdvance := FALSE;

    CASE _eState OF

    E_PlayerState#PS_IDLE:
        bBusy := FALSE;
        wStep := WORD#0;
        dwRequest := DWORD#0;

    E_PlayerState#PS_NEXT_OP:
        (* wStep changes at most once per call: the head checks step + 1 per telegram *)
        IF NOT _bStepSet THEN
            _nOp := _nOp + 1;
            IF _nOp > GVL_Program.N_OPS THEN
                _eState := E_PlayerState#PS_DONE;
            ELSE
                wStep := INT_TO_WORD(_nOp);
                _bStepSet := TRUE;
                _dwMask := GVL_Program.aOps[_nOp].dwZoneMask;
                IF _dwMask <> DWORD#0 THEN
                    dwRequest := _dwMask;           (* same telegram as wStep *)
                    _eState := E_PlayerState#PS_WAIT_GRANT;
                ELSE
                    _rTimer := 0.0;
                    _eState := E_PlayerState#PS_DELAY;
                END_IF
            END_IF
            _bAdvance := TRUE;
        END_IF

    E_PlayerState#PS_WAIT_GRANT:
        IF (dwGrant AND _dwMask) = _dwMask THEN
            _rTimer := 0.0;
            _eState := E_PlayerState#PS_DELAY;
            _bAdvance := TRUE;
        END_IF

    E_PlayerState#PS_DELAY:
        IF _rTimer >= GVL_Program.aOps[_nOp].rDelay_s THEN
            (* Begin the motion of op _nOp *)
            _rT := 0.0;
            _rVel := GVL_Program.aOps[_nOp].rVelScale;
            IF _rVel <= 0.0 THEN
                _rVel := 1.0;
            END_IF
            _bHomeMove := GVL_Program.aOps[_nOp].bBlindHome;
            IF _bHomeMove THEN
                FOR _i := 1 TO 6 DO
                    _arQ0[_i] := _arQ[_i];
                END_FOR
                _rDur := GVL_Program.R_HOME_S;
                _nLast := 0;
            ELSE
                _nWp := GVL_Program.aOps[_nOp].nFirstWp;
                _nLast := GVL_Program.aOps[_nOp].nLastWp;
                IF _nWp < 1 OR _nLast < _nWp OR _nLast > GVL_Program.N_WP THEN
                    _nLast := 0;                    (* no valid trajectory: zero-length move *)
                ELSE
                    (* Start deviation: the trajectory should start at the current pose *)
                    _arQa[1] := GVL_Program.aWp[_nWp].rA1;
                    _arQa[2] := GVL_Program.aWp[_nWp].rA2;
                    _arQa[3] := GVL_Program.aWp[_nWp].rA3;
                    _arQa[4] := GVL_Program.aWp[_nWp].rA4;
                    _arQa[5] := GVL_Program.aWp[_nWp].rA5;
                    _arQa[6] := GVL_Program.aWp[_nWp].rA6;
                    FOR _i := 1 TO 6 DO
                        IF ABS(_arQ[_i] - _arQa[_i]) > GVL_Program.R_START_TOL_DEG THEN
                            wWarningCode := GVL_Program.WARN_START_DEVIATION;
                        END_IF
                    END_FOR
                END_IF
            END_IF
            _eState := E_PlayerState#PS_MOVE;
            _bAdvance := TRUE;
        END_IF

    E_PlayerState#PS_MOVE:
        _bMoveDone := FALSE;
        IF _bHomeMove THEN
            (* Blind joint move: linear in joint space over R_HOME_S *)
            IF _rDur > 0.0 THEN
                _rAlpha := LIMIT(0.0, _rT / _rDur, 1.0);
            ELSE
                _rAlpha := 1.0;
            END_IF
            FOR _i := 1 TO 6 DO
                _arQ[_i] := _arQ0[_i] + _rAlpha * (GVL_Program.arHomeDeg[_i] - _arQ0[_i]);
            END_FOR
            _bMoveDone := _rAlpha >= 1.0;
        ELSIF _nLast < 1 THEN
            _bMoveDone := TRUE;
        ELSE
            (* Trajectory: find the segment [_nWp, _nWp + 1] that contains _rT *)
            WHILE _nWp < _nLast DO
                IF GVL_Program.aWp[_nWp + 1].rT <= _rT THEN
                    _nWp := _nWp + 1;
                ELSE
                    EXIT;
                END_IF
            END_WHILE
            _arQa[1] := GVL_Program.aWp[_nWp].rA1;
            _arQa[2] := GVL_Program.aWp[_nWp].rA2;
            _arQa[3] := GVL_Program.aWp[_nWp].rA3;
            _arQa[4] := GVL_Program.aWp[_nWp].rA4;
            _arQa[5] := GVL_Program.aWp[_nWp].rA5;
            _arQa[6] := GVL_Program.aWp[_nWp].rA6;
            IF _nWp >= _nLast THEN
                FOR _i := 1 TO 6 DO
                    _arQ[_i] := _arQa[_i];
                END_FOR
                _bMoveDone := TRUE;
            ELSE
                _arQb[1] := GVL_Program.aWp[_nWp + 1].rA1;
                _arQb[2] := GVL_Program.aWp[_nWp + 1].rA2;
                _arQb[3] := GVL_Program.aWp[_nWp + 1].rA3;
                _arQb[4] := GVL_Program.aWp[_nWp + 1].rA4;
                _arQb[5] := GVL_Program.aWp[_nWp + 1].rA5;
                _arQb[6] := GVL_Program.aWp[_nWp + 1].rA6;
                _rSpan := GVL_Program.aWp[_nWp + 1].rT - GVL_Program.aWp[_nWp].rT;
                IF _rSpan > 0.0 THEN
                    _rAlpha := LIMIT(0.0, (_rT - GVL_Program.aWp[_nWp].rT) / _rSpan, 1.0);
                ELSE
                    _rAlpha := 1.0;
                END_IF
                FOR _i := 1 TO 6 DO
                    _arQ[_i] := _arQa[_i] + _rAlpha * (_arQb[_i] - _arQa[_i]);
                END_FOR
            END_IF
        END_IF
        IF _bMoveDone THEN
            IF _nOp = 0 THEN
                _eState := E_PlayerState#PS_DONE;   (* HOME_FOLGE finished *)
            ELSE
                _rTimer := 0.0;
                _eState := E_PlayerState#PS_HOLD;
            END_IF
            _bAdvance := TRUE;
        END_IF

    E_PlayerState#PS_HOLD:
        IF _rTimer >= GVL_Program.aOps[_nOp].rHold_s THEN
            IF _dwMask <> DWORD#0 THEN
                dwRequest := DWORD#0;
                _eState := E_PlayerState#PS_WAIT_RELEASE;
            ELSE
                _eState := E_PlayerState#PS_NEXT_OP;
            END_IF
            _bAdvance := TRUE;
        END_IF

    E_PlayerState#PS_WAIT_RELEASE:
        (* 4-phase: the GRANT must drop before the next REQUEST *)
        IF (dwGrant AND _dwMask) = DWORD#0 THEN
            _eState := E_PlayerState#PS_NEXT_OP;
            _bAdvance := TRUE;
        END_IF

    E_PlayerState#PS_DONE:
        bBusy := FALSE;
        bDone := TRUE;
        wStep := WORD#0;
        dwRequest := DWORD#0;
        _eState := E_PlayerState#PS_IDLE;

    E_PlayerState#PS_ERROR:
        bBusy := FALSE;
        bError := TRUE;
        wStep := WORD#0;
        dwRequest := DWORD#0;
        _eState := E_PlayerState#PS_IDLE;

    END_CASE

    IF NOT _bAdvance THEN
        EXIT;
    END_IF
END_FOR

(* ============================================================================
   PUBLISH
   ============================================================================ *)
bAtHome := TRUE;
FOR _i := 1 TO 6 DO
    IF ABS(_arQ[_i] - GVL_Program.arHomeDeg[_i]) > GVL_Program.R_AT_HOME_TOL_DEG THEN
        bAtHome := FALSE;
    END_IF
END_FOR
rA1_deg := _arQ[1];
rA2_deg := _arQ[2];
rA3_deg := _arQ[3];
rA4_deg := _arQ[4];
rA5_deg := _arQ[5];
rA6_deg := _arQ[6];
eState := _eState;
END_FUNCTION_BLOCK
